// TwinCAT 3 PLC project SPS
// ProgramVersion: 3.1.4023.0
// libraries:
//   Tc2_MC2, * (Beckhoff Automation GmbH)
//   Tc2_NCI, * (Beckhoff Automation GmbH)
//   Tc2_PlcInterpolation, * (Beckhoff Automation GmbH)
//   Tc2_Standard, * (Beckhoff Automation GmbH)
//   Tc2_System, * (Beckhoff Automation GmbH)
//   Tc3_Module, * (Beckhoff Automation GmbH)
//   VisuDialogs, * (System)
//   VisuSymbols,3.5.10.0,System
// project tree:
//   DUTs/ E_AxesCmd.TcDUT, E_ButtonState.TcDUT, E_CheckMagazines_New.TcDUT, E_ErrorIDs.TcDUT, E_ErrorSrcs.TcDUT, E_GripperState.TcDUT, E_JobType.TcDUT, E_NC_State.TcDUT, E_NCI_State.TcDUT, E_PortalState.TcDUT, E_PortalState_New.TcDUT, E_ResetHW.TcDUT, E_SetJobState.TcDUT, ST_DeviceState.TcDUT, ST_Channel.TcDUT, ST_Light.TcDUT, ST_Error.TcDUT, ST_PortalJob.TcDUT, ST_PositionCmd.TcDUT, ST_SoftKey.TcDUT
//   / GlobalTextList.TcGTLO, PlcTask.TcTTO, Visualization Manager.TcVMO (not stored), VISU_TASK.TcTTO
//   GVLs/ HMI.TcGVL, GVL_CONST.TcGVL
//   POUs/Aktorik/ FB_AxesEnable.TcPOU, FB_AxisCtrl.TcPOU (excluded from build), FB_Gripper.TcPOU, FB_NciCtrl.TcPOU, FB_SimpleNcControl.TcPOU (excluded from build), FB_VI_Light.TcPOU
//   POUs/ FB_ErrorCollector.TcPOU, FB_IgorCtrl.TcPOU, FB_Portal.TcPOU, MAIN.TcPOU
//   POUs/Safety/ FB_SafeEStop.TcPOU, FB_SafeGroup.TcPOU, FB_SafeMon.TcPOU, FB_SafetyMonitoring.TcPOU
//   POUs/Zeug/ FB_BlockEconomySmart.TcPOU, FB_Error.TcPOU, FB_FuseControl.TcPOU, FB_FuseControl_1.TcPOU, I_NC_Ctrl.TcIO
//   VISUs/ VISU.TcVIS
// real-time tasks:
//   TASK PlcTask: cycle T#10ms, priority 20, ADS port 350
//   TASK PlcTask1: cycle T#10ms, priority 21, ADS port 351
//   TASK VISU_TASK: cycle T#50000us, priority 30, ADS port 352
// motion (NC):
//   TASK NC-Task 1 SAF: cycle T#2ms, priority 4, ADS port 501
//   TASK NC-Task 1 SVB: cycle T#10ms, priority 8, ADS port 511
//   AXIS X (id 1)
//     Dynamic: Acceleration=7500, Deceleration=7500, Jerk=20000, ToleranceBallAuxAxis=20
//     Velo: RefSearch=7.60333333333333, RefSync=7.60333333333333, SlowManual=38.0166666666667, FastManual=750, Fast=760.333333333333, Maximum=760.333
//     TargetPosControl: Range=0.5
//     PEHControl: Enable=true, Time=10
//     OtherSettings: AllowMotionCmdToSlave=true
//     encoder EncType=19
//       EncPara: ScaleFactorNumerator=20, ScaleFactorDenominator=1048576, Offset=150.930252075195, MaxCount=#xffffffff, ReferenceSystem=1
//         SoftEndMinControl: Enable=true, Range=-100
//         SoftEndMaxControl: Enable=true, Range=415
//         TimeComp: TimeCompMode=1
//     drive DrvType=16
//       DrvPara: MaxCount=#xffffffff, DriveControlDWord=#x00020100
//         Analog: VeloReferenz=836.366666666667, VeloScale=32, TorqueSetpointScale=10, ScaleFactorActTorque=0.004
//         TimeComp: TimeCompMode=1, TaskDelayCycles=1
//     controller CtrType=1
//       CtrPara: PriorControlFactor=1
//         PID: PosKp=30
//         Observer: BandWidth=20
//   AXIS Y (id 2)
//     Dynamic: Acceleration=2027.55, Deceleration=2027.55, Jerk=5406.81, ToleranceBallAuxAxis=20
//     Velo: RefSearch=7.60333333333333, RefSync=7.60333333333333, SlowManual=38.0166666666667, FastManual=700, Fast=760.333333333333, Maximum=760.333
//     TargetPosControl: Range=0.5
//     PEHControl: Enable=true, Time=10
//     OtherSettings: AllowMotionCmdToSlave=true
//     encoder EncType=19
//       EncPara: ScaleFactorNumerator=20, ScaleFactorDenominator=1048576, Offset=-52.5408172607422, MaxCount=#xffffffff, ReferenceSystem=1
//         SoftEndMinControl: Enable=true, Range=-2
//         SoftEndMaxControl: Enable=true, Range=300
//         TimeComp: TimeCompMode=1
//     drive DrvType=16
//       DrvPara: MaxCount=#xffffffff, DriveControlDWord=#x00020100
//         Analog: VeloReferenz=836.366666666667, VeloScale=32, TorqueSetpointScale=10, ScaleFactorActTorque=0.1
//         TimeComp: TimeCompMode=1, TaskDelayCycles=1
//     controller CtrType=1
//       CtrPara: PriorControlFactor=1
//         Observer: BandWidth=20
//   AXIS Z (id 3)
//     Dynamic: Acceleration=7500, Deceleration=7500, Jerk=20000, ToleranceBallAuxAxis=20
//     Velo: RefSearch=2.875, RefSync=2.875, SlowManual=14.375, FastManual=200.25, Fast=287.5, Maximum=287.5
//     TargetPosControl: Range=0.5
//     OtherSettings: AllowMotionCmdToSlave=true
//     encoder EncType=19
//       EncPara: ScaleFactorNumerator=5, ScaleFactorDenominator=1048576, Offset=69.1336441040039, Inverse=true, MaxCount=#xffffffff, ReferenceSystem=1
//         SoftEndMinControl: Enable=true
//         SoftEndMaxControl: Enable=true, Range=90
//         TimeComp: TimeCompMode=1
//     drive DrvType=16
//       DrvPara: Inverse=true, MaxCount=#xffffffff, DriveControlDWord=#x00020100
//         Analog: VeloReferenz=316.25, VeloScale=32, TorqueSetpointScale=10, ScaleFactorActTorque=0.1
//         TimeComp: TimeCompMode=1, TaskDelayCycles=1
//     controller CtrType=1
//       CtrPara: PriorControlFactor=1
//         PosDiffControl: Range=0.2
//         PID: PosKp=40
//         Observer: BandWidth=20
// I/O:
//   DEVICE Device, AmsNetId 192.168.1.150.4.1
//     +S1-BC1 (EK1100) [EK1100 EtherCAT Coupler (2A E-Bus)]
//       +S1-SI1 (EL1918) [EL1918, 8Ch. Safety Input 24V, TwinSAFE]
//         modules: Module 2 (FSLOGIC)
//       +S1-SO1 (EL2904) [EL2904, 4 Ch. Safety Output 24V, 0.5A, TwinSAFE]
//         modules: Module 1 (FSOES), Module 2 (DO)
//       +S1-DI1 (EL1804) [EL1804 4Ch. Dig. Input 24V, 3ms]
//       +S1-DI2 (EL1804) [EL1804 4Ch. Dig. Input 24V, 3ms]
//       +S1-DO1 (EL2004) [EL2004 4Ch. Dig. Output 24V, 0.5A]
//       +S1-PM1 (EL7211-9014) [EL7211-9014 1Ch. MDP742 Servo motor output stage with OCT (50V, 4.5A RMS) and STO input]
//       +S1-PM2 (EL7211-9014) [EL7211-9014 1Ch. MDP742 Servo motor output stage with OCT (50V, 4.5A RMS) and STO input]
//       +S1-PM3 (EL7211-9014) [EL7211-9014 1Ch. MDP742 Servo motor output stage with OCT (50V, 4.5A RMS) and STO input]
//       Term 20 (EK1310)
//     Box 21 (VIP2000-1010)
// variable links:
//   Device <-> Device/+S1-BC1 (EK1100)/+S1-SI1 (EL1918)
//     +S1-BC1 (EK1100)/+S1-SO1 (EL2904)/Module 1 (FSOES)/RxPDO/FSOE <-> ConnectionInputs/Message_13 TxPDO
//     +S1-BC1 (EK1100)/+S1-SO1 (EL2904)/Module 1 (FSOES)/TxPDO/FSOE <-> ConnectionOutputs/Message_13 RxPDO
//   NC-Task 1 SAF/Axes/X <-> Device/+S1-BC1 (EK1100)/+S1-PM1 (EL7211-9014)
//     Drive/Inputs/In/nDataIn1 <-> DRV Following error actual value/Following error actual value
//     Drive/Inputs/In/nDataIn3[0] <-> DRV Torque actual value/Torque actual value
//     Drive/Inputs/In/nDcOutputTime <-> InfoData/DcOutputShift
//     Drive/Inputs/In/nState1 <-> DRV Statusword/Statusword
//     Drive/Inputs/In/nState2 <-> DRV Statusword/Statusword @bit 8
//     Drive/Inputs/In/nState4 @bit 1 <-> WcState/InputToggle
//     Drive/Inputs/In/nState4 <-> WcState/WcState
//     Drive/Outputs/Out/nCtrl1 <-> DRV Controlword/Controlword
//     Drive/Outputs/Out/nCtrl2 <-> DRV Controlword/Controlword @bit 8
//     Drive/Outputs/Out/nDataOut1 <-> DRV Target position/Target position
//     Enc/Inputs/In/nDataIn1 <-> FB Position/Position
//     Enc/Inputs/In/nDcInputTime <-> InfoData/DcInputShift
//     Enc/Inputs/In/nState4 @bit 1 <-> WcState/InputToggle
//     Enc/Inputs/In/nState4 <-> WcState/WcState
//   NC-Task 1 SAF/Axes/Y <-> Device/+S1-BC1 (EK1100)/+S1-PM2 (EL7211-9014)
//     Drive/Inputs/In/nDataIn1 <-> DRV Following error actual value/Following error actual value
//     Drive/Inputs/In/nDcOutputTime <-> InfoData/DcOutputShift
//     Drive/Inputs/In/nState1 <-> DRV Statusword/Statusword
//     Drive/Inputs/In/nState2 <-> DRV Statusword/Statusword @bit 8
//     Drive/Inputs/In/nState4 @bit 1 <-> WcState/InputToggle
//     Drive/Inputs/In/nState4 <-> WcState/WcState
//     Drive/Outputs/Out/nCtrl1 <-> DRV Controlword/Controlword
//     Drive/Outputs/Out/nCtrl2 <-> DRV Controlword/Controlword @bit 8
//     Drive/Outputs/Out/nDataOut1 <-> DRV Target position/Target position
//     Enc/Inputs/In/nDataIn1 <-> FB Position/Position
//     Enc/Inputs/In/nDcInputTime <-> InfoData/DcInputShift
//     Enc/Inputs/In/nState4 @bit 1 <-> WcState/InputToggle
//     Enc/Inputs/In/nState4 <-> WcState/WcState
//   NC-Task 1 SAF/Axes/Z <-> Device/+S1-BC1 (EK1100)/+S1-PM3 (EL7211-9014)
//     Drive/Inputs/In/nDataIn1 <-> DRV Following error actual value/Following error actual value
//     Drive/Inputs/In/nDcOutputTime <-> InfoData/DcOutputShift
//     Drive/Inputs/In/nState1 <-> DRV Statusword/Statusword
//     Drive/Inputs/In/nState2 <-> DRV Statusword/Statusword @bit 8
//     Drive/Inputs/In/nState4 @bit 1 <-> WcState/InputToggle
//     Drive/Inputs/In/nState4 <-> WcState/WcState
//     Drive/Outputs/Out/nCtrl1 <-> DRV Controlword/Controlword
//     Drive/Outputs/Out/nCtrl2 <-> DRV Controlword/Controlword @bit 8
//     Drive/Outputs/Out/nDataOut1 <-> DRV Target position/Target position
//     Enc/Inputs/In/nDataIn1 <-> FB Position/Position
//     Enc/Inputs/In/nDcInputTime <-> InfoData/DcInputShift
//     Enc/Inputs/In/nState4 @bit 1 <-> WcState/InputToggle
//     Enc/Inputs/In/nState4 <-> WcState/WcState
//   SPS/SPS Instance <-> Device/+S1-BC1 (EK1100)/+S1-DI1 (EL1804)
//     PlcTask Inputs/MAIN.fbIgorCtrl.fbFuseControl.fbBlockFuse.In <-> Channel 3/Input
//     PlcTask Inputs/MAIN.fbIgorCtrl.fbFuseControl48V.bInFuse <-> Channel 4/Input
//     PlcTask Inputs/MAIN.fbIgorCtrl.fbPortal.fbGripper.bGripperFullClosed <-> Channel 2/Input
//     PlcTask Inputs/MAIN.fbIgorCtrl.fbPortal.fbGripper.bPartSensor <-> Channel 1/Input
//   SPS/SPS Instance <-> Device/+S1-BC1 (EK1100)/+S1-DI2 (EL1804)
//     PlcTask Inputs/MAIN.fbIgorCtrl.fbPortal.bStampZAxis <-> Channel 1/Input
//   SPS/SPS Instance <-> Device/+S1-BC1 (EK1100)/+S1-DO1 (EL2004)
//     PlcTask Outputs/MAIN.fbIgorCtrl.fbFuseControl.fbBlockFuse.Out <-> Channel 3/Output
//     PlcTask Outputs/MAIN.fbIgorCtrl.fbFuseControl48V.bOutFuse <-> Channel 4/Output
//     PlcTask Outputs/MAIN.fbIgorCtrl.fbPortal.fbGripper.bCloseGripper <-> Channel 2/Output
//     PlcTask Outputs/MAIN.fbIgorCtrl.fbPortal.fbGripper.bOpenGripper <-> Channel 1/Output
//   SPS/SPS Instance <-> Device/+S1-BC1 (EK1100)/+S1-PM1 (EL7211-9014)
//     PlcTask Inputs/MAIN.fbIgorCtrl.fbSafetyMonitoring.nDrvInfoData1 <-> DRV Info data 1/Info data 1
//   SPS/SPS Instance <-> Device/+S1-BC1 (EK1100)/+S1-PM2 (EL7211-9014)
//     PlcTask Inputs/MAIN.fbIgorCtrl.fbSafetyMonitoring.nDrvInfoData2 <-> DRV Info data 1/Info data 1
//   SPS/SPS Instance <-> Device/+S1-BC1 (EK1100)/+S1-PM3 (EL7211-9014)
//     PlcTask Inputs/MAIN.fbIgorCtrl.fbSafetyMonitoring.nDrvInfoData3 <-> DRV Info data 1/Info data 1
//   SPS/SPS Instance <-> Device/+S1-BC1 (EK1100)/+S1-SI1 (EL1918)
//     PlcTask Inputs/MAIN.fbIgorCtrl.fbPortal.bSafetyOK <-> StandardInputs/Standard Out Var 20
//     PlcTask Inputs/MAIN.fbIgorCtrl.fbSafetyMonitoring.bEStopButtonOk <-> StandardInputs/Standard Out Var 16
//     PlcTask Inputs/MAIN.fbIgorCtrl.fbSafetyMonitoring.bLightCurtainOk <-> StandardInputs/Standard Out Var 19
//     PlcTask Inputs/MAIN.fbIgorCtrl.fbSafetyMonitoring.fbEStop.nDiag <-> Function Block Info Data/SafetyGruppe.SafetyNetzwerk.FBEstop1 Info Data/Diag
//     PlcTask Inputs/MAIN.fbIgorCtrl.fbSafetyMonitoring.fbEStop.nState <-> Function Block Info Data/SafetyGruppe.SafetyNetzwerk.FBEstop1 Info Data/State
//     PlcTask Inputs/MAIN.fbIgorCtrl.fbSafetyMonitoring.fbGroup.nDiag <-> TwinSAFE Group Info Data/SafetyGruppe Info Data/Diag
//     PlcTask Inputs/MAIN.fbIgorCtrl.fbSafetyMonitoring.fbGroup.nState <-> TwinSAFE Group Info Data/SafetyGruppe Info Data/State
//     PlcTask Inputs/MAIN.fbIgorCtrl.fbSafetyMonitoring.fbMonEStop.nDiag <-> Function Block Info Data/SafetyGruppe.SafetyNetzwerk.FBMon1 Info Data/Diag
//     PlcTask Inputs/MAIN.fbIgorCtrl.fbSafetyMonitoring.fbMonEStop.nState <-> Function Block Info Data/SafetyGruppe.SafetyNetzwerk.FBMon1 Info Data/State
//     PlcTask Inputs/MAIN.fbIgorCtrl.fbSafetyMonitoring.fbMonLightCurtain.nDiag <-> Function Block Info Data/SafetyGruppe.SafetyNetzwerk.FBMon2 Info Data/Diag
//     PlcTask Inputs/MAIN.fbIgorCtrl.fbSafetyMonitoring.fbMonLightCurtain.nState <-> Function Block Info Data/SafetyGruppe.SafetyNetzwerk.FBMon2 Info Data/State
//     PlcTask Inputs/MAIN.fbIgorCtrl.fbSafetyMonitoring.fbMonSafetyGroup.nDiag <-> Function Block Info Data/SafetyGruppe.SafetyNetzwerk.FBMon3 Info Data/Diag
//     PlcTask Inputs/MAIN.fbIgorCtrl.fbSafetyMonitoring.fbMonSafetyGroup.nState <-> Function Block Info Data/SafetyGruppe.SafetyNetzwerk.FBMon3 Info Data/State
//     PlcTask Outputs/MAIN.fbIgorCtrl.fbPortal.bQuitEStop <-> StandardOutputs/Standard In Var 17
//     PlcTask Outputs/MAIN.fbIgorCtrl.fbPortal.bSafetyErrAck <-> StandardOutputs/Standard In Var 23
//     PlcTask Outputs/MAIN.fbIgorCtrl.fbPortal.bSafetyRun <-> StandardOutputs/Standard In Var 22
//     PlcTask Outputs/MAIN.fbIgorCtrl.fbSafetyMonitoring.bCollectEDM <-> StandardOutputs/Standard In Var 24
//   SPS/SPS Instance <-> Device/Box 21 (VIP2000-1010)
//     PlcTask Inputs/MAIN.fbIgorCtrl.fbLight.stDeviceState.Diag <-> Device/Main Inputs/Diag
//     PlcTask Inputs/MAIN.fbIgorCtrl.fbLight.stDeviceState.Error <-> Device/Main Inputs/Error
//     PlcTask Inputs/MAIN.fbIgorCtrl.fbLight.stDeviceState.Ready <-> Device/Main Inputs/Ready
//     PlcTask Inputs/MAIN.fbIgorCtrl.fbLight.stDeviceState.State <-> Device/Main Inputs/Status
//     PlcTask Inputs/MAIN.fbIgorCtrl.fbLight.stDeviceState.SwitchOnCnt <-> Device/Main Inputs/Switch-on counter
//     PlcTask Inputs/MAIN.fbIgorCtrl.fbLight.stDeviceState.Warning <-> Device/Main Inputs/Warning
//     PlcTask Inputs/MAIN.fbIgorCtrl.fbLight.stLight.bLightOn <-> Device/Opmode Continuous Inputs/Light on
//     PlcTask Outputs/MAIN.fbIgorCtrl.fbLight.stLight.bActive <-> Device/Opmode Continuous Outputs/Output
//     PlcTask Outputs/MAIN.fbIgorCtrl.fbLight.stLight.bEnable <-> Device/Main Outputs/Enable
//     PlcTask Outputs/MAIN.fbIgorCtrl.fbLight.stLight.bReset <-> Device/Main Outputs/Reset
//     PlcTask Outputs/MAIN.fbIgorCtrl.fbLight.stLight.channel[1]/bActive <-> Channel Red/ChContinuous Outputs/Active
//     PlcTask Outputs/MAIN.fbIgorCtrl.fbLight.stLight.channel[1]/nBrightness <-> Channel Red/ChContinuous Outputs/Brightness
//     PlcTask Outputs/MAIN.fbIgorCtrl.fbLight.stLight.channel[2]/bActive <-> Channel Blue/ChContinuous Outputs/Active
//     PlcTask Outputs/MAIN.fbIgorCtrl.fbLight.stLight.channel[2]/nBrightness <-> Channel Blue/ChContinuous Outputs/Brightness
//     PlcTask Outputs/MAIN.fbIgorCtrl.fbLight.stLight.channel[3]/bActive <-> Channel Green/ChContinuous Outputs/Active
//     PlcTask Outputs/MAIN.fbIgorCtrl.fbLight.stLight.channel[3]/nBrightness <-> Channel Green/ChContinuous Outputs/Brightness
//     PlcTask Outputs/MAIN.fbIgorCtrl.fbLight.stLight.channel[4]/bActive <-> Channel Orange/ChContinuous Outputs/Active
//     PlcTask Outputs/MAIN.fbIgorCtrl.fbLight.stLight.channel[4]/nBrightness <-> Channel Orange/ChContinuous Outputs/Brightness
//   SPS/SPS Instance <-> NC-Task 1 SAF/Axes/X
//     PlcTask Inputs/MAIN.fbIgorCtrl.fbPortal.aAxis[0].NcToPlc <-> Outputs/ToPlc
//     PlcTask Outputs/MAIN.fbIgorCtrl.fbPortal.aAxis[0].PlcToNc <-> Inputs/FromPlc
//   SPS/SPS Instance <-> NC-Task 1 SAF/Axes/Y
//     PlcTask Inputs/MAIN.fbIgorCtrl.fbPortal.aAxis[1].NcToPlc <-> Outputs/ToPlc
//     PlcTask Outputs/MAIN.fbIgorCtrl.fbPortal.aAxis[1].PlcToNc <-> Inputs/FromPlc
//   SPS/SPS Instance <-> NC-Task 1 SAF/Axes/Z
//     PlcTask Inputs/MAIN.fbIgorCtrl.fbPortal.aAxis[2].NcToPlc <-> Outputs/ToPlc
//     PlcTask Outputs/MAIN.fbIgorCtrl.fbPortal.aAxis[2].PlcToNc <-> Inputs/FromPlc
//   SPS/SPS Instance <-> NC-Task 1 SAF/Interpolation Channel
//     PlcTask Inputs/MAIN.fbIgorCtrl.fbPortal.fbNciCtrl.stItpToPlc <-> Outputs/ToPlc
//     PlcTask Outputs/MAIN.fbIgorCtrl.fbPortal.fbNciCtrl.stPlcToItp <-> Inputs/FromPlc

CONFIGURATION SPS
    RESOURCE PLC ON TwinCAT3
        TASK PlcTask(INTERVAL := T#10ms, PRIORITY := 21);
        TASK VISU_TASK(INTERVAL := T#50000us, PRIORITY := 30);
        PROGRAM MAIN WITH PlcTask : MAIN;
        PROGRAM VisuElems_Visu_Prg WITH VISU_TASK : VisuElems.Visu_Prg;
    END_RESOURCE
END_CONFIGURATION

// ---- DUTs/E_AxesCmd.TcDUT
TYPE E_AxesCmd :
(
	E_AxesCmd_IDLE := 0,
	E_AxesCmd_RESET := 10,
	E_AxesCmd_MOVE_ABS := 20,
	E_AxesCmd_MOVE_REL := 30,
	E_AxesCmd_JOG := 40,
	E_AxesCmd_REFERENCING := 50,
	E_AxesCmd_STOP := 70,
	E_AxesCmd_FINISHED := 80,
	E_AxesCmd_ERROR := 99
);
END_TYPE

// ---- DUTs/E_ButtonState.TcDUT
{attribute 'strict'}
TYPE E_ButtonState :
(
	E_ButtonState_OFF := 0,
	E_ButtonState_ON,
	E_ButtonState_BLINK
);
END_TYPE

// ---- DUTs/E_CheckMagazines_New.TcDUT
{attribute 'qualified_only'}
{attribute 'strict'}
TYPE E_CheckMagazines_New :
(
	eIdle	:= 0,
	eStartNewNCI	:= 1,
	eDebug := 2,
	eWaitForPortal := 3
);
END_TYPE

// ---- DUTs/E_ErrorIDs.TcDUT
{attribute 'qualified_only'}
{attribute 'strict'}
TYPE E_ErrorIDs :
(
	eNoError := 0,
	eUndefinedError := 1,
	eUndefinedState := 2,
	
	eInvalidReference := 21,
	
	eAxisRelease := 31,
	eAbsMove := 32,
	eRelMove := 33,
	eJog := 34,
	eStopAxis := 35,
	eResetAxis := 36,
	eAxesNotReady := 37,
	eAxisError := 38,
	
	eTimeout := 41,
	eInvalidData := 42,
	eReset := 43,
	
	eBuildGroup := 51,
	eClearGroup := 52,
	eFillTable := 53,
	eNotAllowedDriveDown := 54,
	
	eSafetyFbError := 61,
	eCommError := 62,
	eModuleFault := 63,
	eCompareError := 64,
	eEStopPressed := 65,
	eLightCurtain := 66,
	
	eNoStoneInGripper := 71,
	eMagEmpty := 72,
	
	eFuseTripped := 81,
	eFuseOff := 82,
	eFuseOvercurrent := 83,
	
	eClearFieldNoCapacityFound := 90,
	eNoJobsFound := 91,
	eStamp := 92,
	eNoStonesFound := 93,
	
	eCtrlOff := 99
);
END_TYPE

// ---- DUTs/E_ErrorSrcs.TcDUT
{attribute 'qualified_only'}
{attribute 'strict'}
TYPE E_ErrorSrcs :
(
	eNoError := 0,
	ePlc := 1,
	eAxisX := 2,
	eAxisY := 3,
	eAxisZ := 4,
	eAxisGroup := 5,
	eAxisCtrlPtp := 6,
	eAxisCtrlNci := 7,
	eAxisCtrl := 8,
	eGripper := 9,
	eSafety := 10,
	eSafetyGroup := 11,
	eSafetyFb := 12,
	ePortal := 13,
	eFuse := 14
);
END_TYPE

// ---- DUTs/E_GripperState.TcDUT

TYPE E_GripperState :
(
	E_GripperState_INIT := 0,
	E_GripperState_OPENING,
	E_GripperState_OPENED,
	E_GripperState_CLOSING,
	E_GripperState_CLOSED,
	E_GripperState_UNDEFINED
);
END_TYPE

// ---- DUTs/E_JobType.TcDUT
TYPE E_JobType :
(
	E_JobType_MoveStone,
	E_JobType_NewStone,
	E_JobType_RemoveStone
);
END_TYPE

// ---- DUTs/E_NC_State.TcDUT
TYPE E_NC_State :
(
	E_NC_State_INIT := 0,
	E_NC_State_IDLE := 1,
	E_NC_State_RUN := 7,
	E_NC_State_ABORT := 8,
	E_NC_State_ERROR := 9
);
END_TYPE

// ---- DUTs/E_NCI_State.TcDUT
TYPE E_NCI_State :
(
	E_NCI_State_INIT := 0,
	E_NCI_State_IDLE := 1,
	E_NCI_State_BUILD_GROUP := 4,
	E_NCI_State_LOAD_CODE := 5,
	E_NCI_State_FEED_TABLE := 6,
	E_NCI_State_RUN := 7,
	E_NCI_State_ABORT := 8,
	E_NCI_State_CLEAR_GROUP := 9,
	E_NCI_State_ESTOP := 90,
	E_NCI_State_ERROR := 99
);
END_TYPE

// ---- DUTs/E_PortalState.TcDUT
TYPE E_PortalState :
(
	E_PortalState_INIT := 0,
	E_PortalState_IDLE,
	E_PortalState_SET_JOB,
	E_PortalState_MOVE_TO_STONE,
	E_PortalState_TRANSPORT_STONE,
	E_PortalState_WAITGRIPPER_OPEN,
	E_PortalState_WAITGRIPPER_CLOSE,
	E_PortalState_HOME,
	E_PortalState_ESTOP,
	E_PortalState_AFTER_ESTOP,
	E_PortalState_MANUAL_MODE,
	E_PortalState_SCAN_MAGS,
	E_PortalState_ERROR := 99
);
END_TYPE

// ---- DUTs/E_PortalState_New.TcDUT
TYPE E_PortalState_New :
(
	eInit := 0,
	eIdle,
	eSetJob,
	eOpenGripper,
	eCloseGripper,
	eError,
	eMoveToStone,
	eTrspStone,
	eStampTriggered,
	eHome,
	eEStop,
	eAfterEStop,
	eManualMode,
	eDebug
);
END_TYPE

// ---- DUTs/E_ResetHW.TcDUT
{attribute 'qualified_only'}
{attribute 'strict'}
TYPE E_ResetHW :
(
	INIT := 0,
	RESET_HW := 10,
	DONE := 50
);
END_TYPE

// ---- DUTs/E_SetJobState.TcDUT
{attribute 'qualified_only'}
{attribute 'strict'}
TYPE E_SetJobState :
(
	eIdle := 0,
	eAxesNotReady,
	eSelNewStone,
	eSelRemoveStone,
	eCheckAllMagazines,
	eValidateNewStone,
	eValidateRemoveStone
);
END_TYPE

// ---- DUTs/ST_DeviceState.TcDUT
TYPE ST_DeviceState :
STRUCT
	Ready		AT%I*	: BIT;
	Warning		AT%I*	: BIT;
	Error		AT%I*	: BIT;
	Diag		AT%I*	: BIT;
	State		AT%I*	: UDINT;
	SwitchOnCnt	AT%I*	: UDINT;
END_STRUCT
END_TYPE

// ---- DUTs/ST_Channel.TcDUT
TYPE ST_Channel :
STRUCT
	bActive				AT %Q*  : BOOL	 := FALSE;	
	nBrightness			AT %Q*	: UINT	 := 100; 
END_STRUCT
END_TYPE

// ---- DUTs/ST_Light.TcDUT
TYPE ST_Light :
STRUCT
	bEnable					AT %Q* 	: BOOL := TRUE;				// Global enable of light
	bReset					AT %Q*	: BOOL := FALSE;			// Reset light
	bActive					AT %Q*  : BOOL	 := FALSE;			// General activation of the light, depends on the chanels
	bLightOn				AT %I*	: BOOL;						// Light is activated
	channel					AT %Q*  : ARRAY[1..4] OF ST_Channel; // 1: IR, 2: blue, 3: green, 4: orange
	nTemperature			AT %I*	: SINT;						// temperature channel
END_STRUCT
END_TYPE

// ---- DUTs/ST_Error.TcDUT
TYPE ST_Error :
STRUCT
	nSource:		UDINT;
	nType:			UDINT;
	sMsg:			STRING(80);
END_STRUCT
END_TYPE

// ---- DUTs/ST_PortalJob.TcDUT
TYPE ST_PortalJob :
STRUCT
	nJobID:			UDINT; //Job Nummer
	eJobType:		E_JobType;  //Neuer Stein von Stapel oder Stein auf Brett oder Stein entfernen
	fStartPosX:		LREAL; //Startposition x in mm
	fStartPosY:		LREAL; //Startposition y in mm
	fDestPosX:		LREAL; //Zielposition x in mm
	fDestPosY:		LREAL; //Zielposition y in mm
	bBlack:			BOOL; //entscheidet über Lagerposition
END_STRUCT
END_TYPE

// ---- DUTs/ST_PositionCmd.TcDUT
TYPE ST_PositionCmd :
STRUCT
	nNo:	UDINT;
	fPosX:	LREAL;
	fPosY:	LREAL;
	fPosZ:	LREAL;
	fVelo:	LREAL;
	bExact:	BOOL;
END_STRUCT
END_TYPE

// ---- DUTs/ST_SoftKey.TcDUT
TYPE ST_SoftKey :
STRUCT
	bIsPressed:	BOOL;
	eState:		E_ButtonState;
END_STRUCT
END_TYPE

// ---- GVLs/HMI.TcGVL
{attribute 'qualified_only'}
VAR_GLOBAL	
//TO HMI
	bErrorChange:		BOOL;
	aErrors:			ARRAY [0..MAX_ERRORS - 1] OF ST_Error;
	nNumberErrors:		UINT;
	bSafetyOK:			BOOL;
	bPortalBusy:		BOOL;
	bInManual:			BOOL;
	bGripperOpen:		BOOL;
	bGripperClosed:		BOOL;
	bHandInPortal:		BOOL; 
	
//FROM HMI
	bQuit:				BOOL;
	
	bSetJob:			BOOL;
	stJob:				ST_PortalJob;
	stLastJob:			ST_PortalJob;
     	
	bReqManualCtrl:		BOOL := TRUE;
	bOpenGripper:		BOOL;
	bCloseGripper:		BOOL;
	bSafetyRun:			BOOL;
	
	bLightOn:			BOOL;
	bLightWin: 			BOOL;
	bLightLose:			BOOL;
	
	bLightParty: 		BOOL;
	
	bAllJobsSend: 		BOOL; 
	
//TO AND FROM HMI
	stSoftKeyCtrlOn:	ST_SoftKey;
	stSoftKeyCtrlOff:	ST_SoftKey;
	stSoftKeyAutoOn:	ST_SoftKey;
	stSoftKeyAutoOff:	ST_SoftKey;
	stSoftKeyQuit:		ST_SoftKey;

//system
	fbErrorCollector:	FB_ErrorCollector;
	
//parameters
	fAxesOverride:		LREAL := 100.0;
	fAxesOverrideMan:	LREAL := 20.0;
	
	fPortalPosIdleX:	LREAL := -20;
	fPortalPosIdleY:	LREAL := 0;
	fPortalPosIdleZ:	LREAL := 50;

	fScreenPosOffsetX:	LREAL := 0;
	fScreenPosOffsetY:	LREAL := 0;
END_VAR

// ---- GVLs/GVL_CONST.TcGVL
VAR_GLOBAL CONSTANT	
	STONE_POS_FIELD_Z:	LREAL := 1;
	MIN_MOVE_HEIGHT_Z:	LREAL := 40; //beachte: Stäbe von Magazin ca. 35 mm -> nicht unter 40 stellen!
	STONE_HEIGHT:		LREAL := 8; //Steinhöhe in mm -> für Positionen in Magazin
	
	MAX_JOB_COUNT:		USINT := 30;
	MAX_ERRORS:			USINT := 55;
	
	X:					USINT := 0;
	Y:					USINT := 1;
	Z:					USINT := 2;
	
	MAGAZINE_NUMBER:	USINT := 6; //Anzahl Magazine
	MAGAZINE_CAPACITY:	USINT := 4;	//Anzahl Positionen pro Magazin	
	
(******Stapel für Spielsteine******)
	STACK_POS_X:			LREAL := -97.2; 
	STACK_1_POS_Y:			LREAL := 52.6;	
	STACK_2_POS_Y:			LREAL := STACK_1_POS_Y + 28;
	STACK_3_POS_Y:			LREAL := STACK_2_POS_Y + 28;
	STACK_4_POS_Y:			LREAL := STACK_3_POS_Y + 94;
	STACK_5_POS_Y:			LREAL := STACK_4_POS_Y + 28;
	STACK_6_POS_Y:			LREAL := STACK_5_POS_Y + 28;//258.6
	STACK_POS_Z_BASE:		LREAL := 3;
	STACK_POS_Z_BASE_REMOVE:LREAL := 8;
	
(******Positionen Magazin-Scan******)
	STACK_SCAN_POS_X:		LREAL := -59;
	STACK_1_SCAN_POS_Y:		LREAL := STACK_1_POS_Y + 33.8;
	STACK_2_SCAN_POS_Y:		LREAL := STACK_2_POS_Y + 33.8;
	STACK_3_SCAN_POS_Y:		LREAL := STACK_3_POS_Y + 33.8;
	STACK_4_SCAN_POS_Y:		LREAL := STACK_4_POS_Y + 33.8;
	STACK_5_SCAN_POS_Y:		LREAL := STACK_5_POS_Y + 33.8;
	STACK_6_SCAN_POS_Y:		LREAL := STACK_6_POS_Y + 33.8;
	STACK_SCAN_POS_Z_BASE:	LREAL := 8.5;
	
END_VAR

// ---- POUs/Zeug/I_NC_Ctrl.TcIO
INTERFACE I_NC_Ctrl

METHOD M_AxisRef
VAR_INPUT
	rX:		REFERENCE TO AXIS_REF;
	rY:		REFERENCE TO AXIS_REF;
	rZ:		REFERENCE TO AXIS_REF;
END_VAR
END_METHOD

METHOD M_CancleJob
VAR_INPUT
END_VAR
END_METHOD

METHOD M_Cyclic
VAR_INPUT
END_VAR
END_METHOD

METHOD M_NewJob
VAR_INPUT
	fTargetPosX:	LREAL;
	fTargetPosY:	LREAL;
	fTargetPosZ:	LREAL;
END_VAR
END_METHOD

PROPERTY P_bInductiveSensor : BOOL
SET
END_SET
END_PROPERTY

PROPERTY P_Busy : BOOL
GET
END_GET
END_PROPERTY

PROPERTY P_Enable : BOOL
SET
END_SET
END_PROPERTY

PROPERTY P_ErrID : E_ErrorIDs
GET
END_GET
END_PROPERTY

PROPERTY P_Error : BOOL
GET
END_GET
END_PROPERTY

PROPERTY P_ErrSrc : E_ErrorSrcs
GET
END_GET
END_PROPERTY

PROPERTY P_ReadyForJob : BOOL
GET
END_GET
END_PROPERTY

PROPERTY P_Reset : BOOL
SET
END_SET
END_PROPERTY

END_INTERFACE

// ---- POUs/MAIN.TcPOU
PROGRAM MAIN
VAR
	fbIgorCtrl:			FB_IgorCtrl;
END_VAR

fbIgorCtrl();

END_PROGRAM

// ---- POUs/FB_IgorCtrl.TcPOU
FUNCTION_BLOCK FB_IgorCtrl
VAR_INPUT
END_VAR
VAR_OUTPUT
	fbError:	FB_Error;
END_VAR
VAR
	fbPortal:			FB_Portal;
	fbSafetyMonitoring:	FB_SafetyMonitoring;
	fbFuseControl:		FB_FuseControl;
	fbFuseControl48V: 	FB_FuseControl_1;
	fbLight			:	FB_VI_Light;
END_VAR

VAR
	fbBlinkTimer1		: TON;
	fbBlinkTimer2		: TON;
	fbTimer				: TON;
	fbRS				: RS;
	nCntParty			: UINT;
	rTrig1				: R_TRIG;
	rTrig2				: R_TRIG;
	
	nRed				: UINT;
	nGreen				: UINT;
	nBlue				: UINT;
END_VAR

A_HmiComm();

fbSafetyMonitoring();

fbFuseControl();
fbFuseControl48V(bResetChannels := HMI.bQuit);


fbPortal(
	bFuseOk := NOT fbFuseControl.fbError.bError,
	bFuse48VOk := NOT fbFuseControl.fbError.bError,
	bManualMode:= HMI.bReqManualCtrl, 
	stNewJob:= HMI.stJob, 
	bImportJob:= HMI.bSetJob,
	bQuit:= HMI.bQuit OR fbPortal.bQuit,//kann quit nicht false setzen
	bSafetyRun := HMI.bSafetyRun,
	bSafetyOK=> HMI.bSafetyOK, 
	bBusy=> HMI.bPortalBusy,
	fbError=> );

HMI.bGripperClosed := fbPortal.fbGripper.bGripperClosed;
HMI.bGripperOpen := fbPortal.fbGripper.bGripperOpen;

IF NOT HMI.bSafetyRun AND NOT fbError.bError THEN
	fbError.M_Set(1, 'Steuerung ausgeschaltet', 0, E_ErrorIDs.eCtrlOff, E_ErrorSrcs.ePlc);
ELSIF HMI.bSafetyRun AND fbError.bError THEN
	fbError.M_Reset();
END_IF

//Set trigger white light
IF HMI.bLightOn THEN
	HMI.bLightWin := FALSE;
	HMI.bLightLose := FALSE;
	fbLight(bLightOn:= HMI.bLightOn);
	fbLight.bLightOn := FALSE;
	fbLight.SetIRGB(255, 255, 255, 255, 100);
ELSIF NOT HMI.bLightWin AND NOT HMI.bLightLose THEN
	fbLight(bLightOn:= HMI.bLightOn);
END_IF

//Set light for win
IF HMI.bLightWin AND NOT HMI.bLightLose AND NOT HMI.bLightOn THEN
	fbTimer(IN := TRUE, PT := T#3S);
	fbRS(SET := TRUE, RESET1 := fbTimer.Q);
	
	fbBlinkTimer1(IN := fbRS.Q1 AND NOT fbBlinkTimer2.Q, PT := T#0.5S, Q => fbLight.bLightOn);
	fbBlinkTimer2(IN := fbBlinkTimer1.Q, PT := T#0.5S);
	fbLight.SetIRGB(0, 0, 255, 0, 50);
	
	IF fbTimer.Q THEN
		HMI.bLightWin := FALSE;
		fbLight.bLightOn := FALSE;
		fbTimer(IN := FALSE);
		fbRS(SET := FALSE, RESET1 := TRUE);
	END_IF
	
	fbLight();
ELSE
	fbRS(SET := FALSE, RESET1 := FALSE);
END_IF

//set light for lose
IF HMI.bLightLose AND NOT HMI.bLightWin AND NOT HMI.bLightOn THEN
	fbTimer(IN := TRUE, PT := T#3S);
	fbRS(SET := TRUE, RESET1 := fbTimer.Q);
	
	fbBlinkTimer1(IN := fbRS.Q1 AND NOT fbBlinkTimer2.Q, PT := T#0.5S, Q => fbLight.bLightOn);
	fbBlinkTimer2(IN := fbBlinkTimer1.Q, PT := T#0.5S);
	fbLight.SetIRGB(0, 255, 0, 0, 50);
	
	IF fbTimer.Q THEN
		HMI.bLightLose := FALSE;
		fbLight.bLightOn := FALSE;
		fbTimer(IN := FALSE);
		fbRS(SET := FALSE, RESET1 := TRUE);
	END_IF
	
	fbLight();
ELSE
	fbRS(SET := FALSE, RESET1 := FALSE);
END_IF

//Party-Modus
IF HMI.bLightParty THEN
	fbTimer(IN := TRUE, PT := T#30S);
	fbRS(SET := TRUE, RESET1 := fbTimer.Q);
	
	fbBlinkTimer1(IN := fbRS.Q1 AND NOT fbBlinkTimer2.Q, PT := T#0.4S, Q => );
	fbBlinkTimer2(IN := fbBlinkTimer1.Q, PT := T#0.2S);
	fbLight.bLightOn := NOT fbBlinkTimer1.Q;
	IF rTrig1.Q OR rTrig2.Q THEN
		nCntParty := nCntParty + 1;
	END_IF
	
	CASE nCntParty OF 
		0: fbLight.SetIRGB(0, 255, 0, 0, 25);
		1: fbLight.SetIRGB(0, 255, 30, 0, 25);
		2: fbLight.SetIRGB(0, 255, 255, 0, 25);
		3: fbLight.SetIRGB(0, 180, 255, 0, 25);
		4: fbLight.SetIRGB(0, 0, 255, 0, 25);
		5: fbLight.SetIRGB(0, 0, 255, 150, 25);
		6: fbLight.SetIRGB(0, 0, 255, 255, 25);
		7: fbLight.SetIRGB(0, 0, 120, 255, 25);
		8: fbLight.SetIRGB(0, 0, 0, 255, 25);
		9: fbLight.SetIRGB(0, 120, 0, 255, 25);
		10: fbLight.SetIRGB(0, 255, 0, 120, 25); nCntParty := 0;
	END_CASE

	IF fbTimer.Q THEN
		HMI.bLightParty := FALSE;
		nCntParty := 0;
		fbLight.bLightOn := FALSE;
		fbTimer(IN := FALSE);
		fbRS(SET := FALSE, RESET1 := TRUE);
	END_IF
	
	rTrig1(CLK := fbBlinkTimer1.Q);
	rTrig2(CLK := fbBlinkTimer2.Q);
	fbLight();
ELSE
	fbRS(SET := FALSE, RESET1 := FALSE);
END_IF

ACTION A_HmiComm:
IF HMI.stSoftKeyCtrlOn.bIsPressed THEN
	HMI.bSafetyRun := TRUE;
END_IF
IF HMI.stSoftKeyCtrlOff.bIsPressed THEN
	HMI.bSafetyRun := FALSE;
END_IF
IF HMI.stSoftKeyAutoOn.bIsPressed THEN
	HMI.bReqManualCtrl := FALSE;
END_IF
IF HMI.stSoftKeyAutoOff.bIsPressed THEN
	HMI.bReqManualCtrl := TRUE;
END_IF

HMI.bInManual := MAIN.fbIgorCtrl.fbPortal.ePortalState = E_PortalState_New.eManualMode;

HMI.bHandInPortal := NOT MAIN.fbIgorCtrl.fbSafetyMonitoring.bLightCurtainOk;

HMI.bQuit := HMI.stSoftKeyQuit.bIsPressed;

IF HMI.bSafetyOK THEN
	HMI.stSoftKeyCtrlOn.eState := E_ButtonState_ON;
	HMI.stSoftKeyCtrlOff.eState := E_ButtonState_OFF;
	
	IF HMI.bReqManualCtrl THEN
		IF Main.fbIgorCtrl.fbPortal.ePortalState <> E_PortalState_New.eManualMode THEN
			HMI.stSoftKeyAutoOn.eState := E_ButtonState_BLINK;
			HMI.stSoftKeyAutoOff.eState := E_ButtonState_OFF;
		ELSE
			HMI.stSoftKeyAutoOn.eState := E_ButtonState_OFF;
			HMI.stSoftKeyAutoOff.eState := E_ButtonState_ON;
		END_IF
	ELSE
		IF HMI.nNumberErrors = 0 THEN
			HMI.stSoftKeyAutoOn.eState := E_ButtonState_ON;
			HMI.stSoftKeyAutoOff.eState := E_ButtonState_OFF;
		ELSE
			HMI.stSoftKeyAutoOn.eState := E_ButtonState_OFF;
			HMI.stSoftKeyAutoOff.eState := E_ButtonState_BLINK;
		END_IF
	END_IF
	
	IF HMI.nNumberErrors > 0 THEN
		HMI.stSoftKeyQuit.eState := E_ButtonState_BLINK;
	ELSE
		HMI.stSoftKeyQuit.eState := E_ButtonState_OFF;
	END_IF
ELSE
	HMI.stSoftKeyAutoOn.eState := E_ButtonState_OFF;
	HMI.stSoftKeyAutoOff.eState := E_ButtonState_ON;
	IF HMI.bSafetyRun THEN
		HMI.stSoftKeyCtrlOn.eState := E_ButtonState_BLINK;
		HMI.stSoftKeyCtrlOff.eState := E_ButtonState_OFF;
		HMI.stSoftKeyQuit.eState := E_ButtonState_BLINK;
	ELSE
		HMI.stSoftKeyCtrlOn.eState := E_ButtonState_OFF;
		HMI.stSoftKeyCtrlOff.eState := E_ButtonState_ON;
		HMI.stSoftKeyQuit.eState := E_ButtonState_OFF;
	END_IF
END_IF
END_ACTION

END_FUNCTION_BLOCK

// ---- POUs/Zeug/FB_Error.TcPOU
{attribute 'reflection'}
FUNCTION_BLOCK FB_Error
VAR_OUTPUT
	bError:		BOOL;
	nErrorID:	UDINT;
	eErrorID:	E_ErrorIDs;
	eErrorSrc:	E_ErrorSrcs;
	sErrorMsg:	STRING(128);
	nState:		INT; //State in dem der Error aufgetreten ist
	
	//{attribute 'instance-path'}
	//{attribute 'no_init'}
	//sSource:	STRING;
END_VAR

METHOD M_Reset
VAR_INPUT
END_VAR
IF bError THEN
	HMI.fbErrorCollector.M_QuitError(eErrorID, eErrorSrc);
	MEMSET(ADR(THIS^), 0, SIZEOF(THIS^));
END_IF
END_METHOD

METHOD M_Set
VAR_INPUT
	nID:	UDINT;
	sMsg:	STRING;
	nState:	INT; //State in dem der Error aufgetreten ist
	eID:	E_ErrorIDs;
	eSrc:	E_ErrorSrcs;
END_VAR
VAR_INST
	
END_VAR
IF NOT bError THEN
	bError := TRUE;
	nErrorID := nID;
	sErrorMsg := sMsg;
	THIS^.nState := nState;
	eErrorID := eID;
	eErrorSrc := eSrc;
	HMI.fbErrorCollector.M_NewError(eID, eSrc, sMsg);
END_IF
END_METHOD

END_FUNCTION_BLOCK

// ---- POUs/FB_Portal.TcPOU
FUNCTION_BLOCK FB_Portal
VAR_INPUT
	bManualMode:			BOOL;	                    	
	stNewJob:				ST_PortalJob;
	bImportJob:				BOOL;
	bQuit:					BOOL;
	bFuseOk:				BOOL;
	bFuse48VOk:				BOOL;
	bSafetyRun AT %Q*:		BOOL;
END_VAR
VAR CONSTANT	
END_VAR                 	
VAR_OUTPUT          		
	bBusy:					BOOL;
	fbError:				FB_Error;
	                    	
	//Safety            	
	bSafetyOK AT %I*:		BOOL := TRUE;
END_VAR             		
VAR                     
	//Safety            	
	bQuitEStop AT %Q*:		BOOL;
	bSafetyErrAck AT %Q*:	BOOL;
	
	//Sensor Stempeln		
	bStampZAxis				AT %I*	: BOOL;
	rTrigStamp:				R_TRIG;
	bStampReset: 			BOOL;
	
	fbRTrigSafety:			R_TRIG;
	                    	
	ePortalState:			E_PortalState_New;
	eTargetPortalState: 	E_PortalState_New;
	                    	
	fbGripper:				FB_Gripper := (bEnable := TRUE);
  
	aAxis:					ARRAY [X..Z] OF AXIS_REF;
	fbAxesEnable:			FB_AxesEnable;
	fbResetAxis:			MC_Reset; 
	                    	
	ipNcCtrl:				I_NC_Ctrl;
	fbNciCtrl:				FB_NciCtrl;
	                    	
	bMagazineTrack:			BOOL; //Anzahl steine in Magazinen bekannt? false wenn Spieler eingreift oder nicht initialisiert
	                    	
	stActJob:				ST_PortalJob;
	aJobBuffer:				ARRAY [0..MAX_JOB_COUNT - 1] OF ST_PortalJob;
	nJobCount:				USINT;
	i, k:					USINT;
	                    	
	aMagCounter:			ARRAY [0..MAGAZINE_NUMBER-1] OF USINT; //Anzahl Steine in Magazinen
	aMagSkipCheck:			ARRAY [0..MAGAZINE_NUMBER-1] OF BOOL;
	aMagYPositions:			ARRAY [0..MAGAZINE_NUMBER-1] OF LREAL; //Mitte Y
	aMagYScanPositions:		ARRAY [0..MAGAZINE_NUMBER-1] OF LREAL;
	fStonePosZFromMag:		LREAL; //berechnete Z pos für Stein aus Magazin
	nMag:					INT;
	nSelectedMag:			INT;
	nPosInMag:				USINT;
	bValidateStonePos:		BOOL;
	nValidationValue:		INT;
	bLastJobBlack:			BOOL;
	
//MAG Check
	nStonesInMag:				INT := MAGAZINE_CAPACITY;
	bWaitPortal, bCheck:		BOOL;
	bCheckedAllMag: 	BOOL;
	nNumChecked:				INT;
	rTrigCheck:			R_TRIG;
//New
	nCntActiveJobs		: SINT;
	nCntRemoveStones	: SINT;
	eCheckMagState		: E_CheckMagazines_New;
	nStonesInMagazin	: USINT := MAGAZINE_CAPACITY;
	
	bAllJobsReceived	: BOOL;
	
	nStateJobSelect		: INT;
	
	bReady				: BOOL;
	
	fTrigNCIDone		: F_TRIG;
	
	fSetJobHeight	: LREAL;
	
	bNCIJobStarted : BOOL;
	
	eSetJobState	: E_SetJobState;
END_VAR

IF ipNcCtrl <> 0 THEN
	A_Cycle();
ELSIF ePortalState <> E_PortalState_INIT THEN
	fbError.M_Set(1, 'Interface nicht referenziert', ePortalState, E_ErrorIDs.eInvalidReference, E_ErrorSrcs.ePlc);
	RETURN;
END_IF
fTrigNCIDone(CLK := fbNciCtrl.P_Busy);

CASE ePortalState OF
	E_PortalState_New.eInit:
		A_Init();
		ePortalState := E_PortalState_New.eIdle;
		
	E_PortalState_New.eIdle:
		IF NOT bManualMode THEN
			IF aJobBuffer[0].nJobID <> 0 THEN
				fbAxesEnable.M_EnableAxes();
				IF fbGripper.bGripperOpen THEN
					IF HMI.bAllJobsSend THEN	
						nValidationValue := 0;	//TODO: entfernen wenn eSetJobState verwendet
						bReady := FALSE;
						nNumChecked := 0;		//TODO: entfernen wenn eSetJobState verwendet
						nStateJobSelect := 0;
						ePortalState := E_PortalState_New.eSetJob;
					END_IF
				ELSE
					eTargetPortalState := E_PortalState_New.eIdle;
					ePortalState := E_PortalState_New.eOpenGripper;
				END_IF
			END_IF
		ELSE	//Handbetrieb
			ipNcCtrl.P_Enable := FALSE;
			fbAxesEnable.M_EnableAxes();
			ePortalState := E_PortalState_New.eManualMode;
		END_IF
	
	E_PortalState_New.eOpenGripper:
		fbGripper(bEnable := TRUE, bOpen := TRUE, bClose := FALSE);
		IF NOT fbGripper.bBusy AND fbGripper.bGripperOpen THEN
			IF eTargetPortalState = E_PortalState_New.eIdle THEN
				fbGripper(bOpen := FALSE);
				ePortalState := eTargetPortalState;	
			ELSE
				IF NOT fbGripper.fbError.bError THEN
					IF stActJob.nJobID <> 0 THEN	//aktuellen Auftrag umgesetzt
						IF stActJob.eJobType = E_JobType.E_JobType_RemoveStone AND nCntActiveJobs = 1 THEN
							aMagCounter[nSelectedMag] := aMagCounter[nSelectedMag] + nCntRemoveStones;
							nCntRemoveStones := 0;
						END_IF
						nCntActiveJobs := nCntActiveJobs - 1;
						HMI.stLastJob := stActJob;
						A_DequeueJob();
						IF nCntActiveJobs <= 0 THEN
							bReady := FALSE;
						END_IF
					ELSE
						bReady := FALSE;
					END_IF
					IF nJobCount = 0 THEN
						ipNcCtrl.M_NewJob(HMI.fPortalPosIdleX, HMI.fPortalPosIdleY, HMI.fPortalPosIdleZ); //Auftrag zu Home-Pos
						ePortalState := E_PortalState_New.eHome;
					ELSE
						ePortalState := E_PortalState_New.eSetJob;	
					END_IF			
				ELSE
					fbError := fbGripper.fbError;
					ePortalState := E_PortalState_New.eError;		
				END_IF
			END_IF
		END_IF
		
	E_PortalState_New.eSetJob:
		HMI.bAllJobsSend := FALSE;
		IF bReady THEN
			//Weiterer Auftrag in Auftragsreihenfolge
			IF nCntActiveJobs >= 1 AND aJobBuffer[0].eJobType = E_JobType.E_JobType_NewStone THEN 
				aJobBuffer[0].fStartPosX := stActJob.fDestPosX;
				aJobBuffer[0].fStartPosY := stActJob.fDestPosY;
				stActJob := aJobBuffer[0];
				
				eTargetPortalState := E_PortalState_New.eMoveToStone;
				ePortalState := E_PortalState_New.eDebug;
				fSetJobHeight := STONE_POS_FIELD_Z + STONE_HEIGHT;
				
				//ipNcCtrl.M_NewJob(stActJob.fStartPosX, stActJob.fStartPosY, STONE_POS_FIELD_Z + STONE_HEIGHT);
				//ePortalState := E_PortalState_New.eMoveToStone;
			//Weiterer Auftrag in Auftragsreihenfolge
			ELSIF nCntActiveJobs >= 1 AND aJobBuffer[0].eJobType = E_JobType.E_JobType_RemoveStone THEN 
				aJobBuffer[0].fStartPosX := stActJob.fDestPosX;
				aJobBuffer[0].fStartPosY := stActJob.fDestPosY;
				stActJob := aJobBuffer[0];
				
				eTargetPortalState := E_PortalState_New.eMoveToStone;
				ePortalState := E_PortalState_New.eDebug;
				fSetJobHeight := STONE_POS_FIELD_Z; 
				
				//ipNcCtrl.M_NewJob(stActJob.fStartPosX, stActJob.fStartPosY, STONE_POS_FIELD_Z);
				//ePortalState := E_PortalState_New.eMoveToStone;
			END_IF
		ELSE
			nStateJobSelect := M_SetJob_New();
			CASE nStateJobSelect OF
				-1: ePortalState := E_PortalState_New.eEStop;
				0: bReady := FALSE;
				1: bReady := TRUE;
					//Mehr als ein gleichzeitiger Auftrag (NewStone)
					IF nCntActiveJobs >= 1 AND aJobBuffer[0].eJobType = E_JobType.E_JobType_NewStone THEN		
						stActJob := aJobBuffer[0];
						//ipNcCtrl.M_NewJob(stActJob.fStartPosX, stActJob.fStartPosY, fStonePosZFromMag);
						//ePortalState := E_PortalState_New.eMoveToStone;
						fSetJobHeight := fStonePosZFromMag;
						eTargetPortalState := E_PortalState_New.eMoveToStone;
						ePortalState := E_PortalState_New.eDebug;
					//Mehr als ein gleichzeitiger Auftrag (RemoveStone)
					ELSIF nCntActiveJobs >= 1 AND aJobBuffer[0].eJobType = E_JobType.E_JobType_RemoveStone THEN
						stActJob := aJobBuffer[0];
						//ipNcCtrl.M_NewJob(stActJob.fStartPosX, stActJob.fStartPosY, STONE_POS_FIELD_Z);
						//ePortalState := e_PortalState_New.eMoveToStone;
						fSetJobHeight := STONE_POS_FIELD_Z;
						eTargetPortalState := E_PortalState_New.eMoveToStone;
						ePortalState := E_PortalState_New.eDebug;
					//Normaler MoveStone-Auftrag
					ELSIF nCntActiveJobs <= -1 THEN	
						stActJob := aJobBuffer[0];
						ipNcCtrl.M_NewJob(stActJob.fStartPosX, stActJob.fStartPosY, STONE_POS_FIELD_Z);
						ePortalState := E_PortalState_New.eMoveToStone;
					ELSE
						ipNcCtrl.M_NewJob(HMI.fPortalPosIdleX, HMI.fPortalPosIdleY, HMI.fPortalPosIdleZ);
						ePortalState := E_PortalState_New.eHome; //oder Error???
					END_IF
			END_CASE
		END_IF
			
	E_PortalState_New.eDebug:
		IF NOT ipNcCtrl.P_Busy THEN
			ipNcCtrl.M_NewJob(stActJob.fStartPosX, stActJob.fStartPosY, fSetJobHeight);
			ePortalState := eTargetPortalState;
		END_IF
	
	E_PortalState_New.eMoveToStone:
		IF NOT ipNcCtrl.P_Busy THEN 				//Warten bis Position erreicht
			IF ipNcCtrl.P_Error THEN				//Error
				fbError.M_Set(1, 'Achsenfehler', ePortalState, eID := ipNcCtrl.P_ErrID, eSrc := ipNcCtrl.P_ErrSrc);
				ePortalState := E_PortalState_New.eError;
			ELSE
				eTargetPortalState := E_PortalState_New.eTrspStone;
				ePortalState := E_PortalState_New.eCloseGripper;
			END_IF 
		END_IF
		
	E_PortalState_New.eCloseGripper:
		fbGripper(bEnable := TRUE, bClose := TRUE, bOpen := FALSE);
		IF NOT fbGripper.bBusy AND fbGripper.bGripperClosed THEN
			IF NOT fbGripper.fbError.bError THEN
				fbGripper(bClose := FALSE);
				IF fbGripper.bStoneInGripper THEN //Stein von Teilesensor erkannt
					IF stActJob.eJobType = E_JobType_NewStone THEN //Stein aus Magazin entnommen
						IF NOT bStampReset THEN
							aMagCounter[nSelectedMag] := aMagCounter[nSelectedMag] - 1;
						ELSE
							bStampReset := FALSE;
						END_IF
						ipNcCtrl.M_NewJob(stActJob.fDestPosX, stActJob.fDestPosY, STONE_POS_FIELD_Z); 
					ELSIF stActJob.eJobType = E_JobType.E_JobType_RemoveStone AND nCntActiveJobs > 1 AND aJobBuffer[1].fStartPosX <> 0 AND aJobBuffer[1].fStartPosY <> 0 THEN
						stActJob.fDestPosX := aJobBuffer[1].fStartPosX;
						stActJob.fDestPosY := aJobBuffer[1].fStartPosY;
						ipNcCtrl.M_NewJob(stActJob.fDestPosX, stActJob.fDestPosY, STONE_POS_FIELD_Z + STONE_HEIGHT);
					ELSIF (stActJob.eJobType = E_JobType.E_JobType_RemoveStone AND nCntActiveJobs = 1) OR (stActJob.eJobType = E_JobType.E_JobType_RemoveStone AND aJobBuffer[1].fStartPosX <> 0 AND aJobBuffer[1].fStartPosY <> 0) THEN
						stActJob.fDestPosX := STACK_POS_X;
						stActJob.fDestPosY := aMagYPositions[nSelectedMag];
						ipNcCtrl.M_NewJob(stActJob.fDestPosX, stActJob.fDestPosY, STACK_POS_Z_BASE_REMOVE + (nPosInMag-1)*STONE_HEIGHT);
					ELSIF stActJob.eJobType =  E_JobType.E_JobType_MoveStone THEN
						ipNcCtrl.M_NewJob(stActJob.fDestPosX, stActJob.fDestPosY, STONE_POS_FIELD_Z); 
					END_IF
					ePortalState := eTargetPortalState;					
				ELSE
					fbError.M_Set(1804, 'Keinen Stein gegriffen!', ePortalState, eID := E_ErrorIDs.eNoStoneInGripper, eSrc := E_ErrorSrcs.eGripper);
					fbGripper(bOpen := TRUE);
					IF aJobBuffer[0].nJobID = 0 THEN
						ePortalState := E_PortalState_New.eIdle;
					ELSE
						bReady := FALSE;
						ePortalState := E_PortalState_New.eSetJob;
					END_IF
				END_IF
			ELSE
				fbError := fbGripper.fbError;
				ePortalState := E_PortalState_New.eError;
			END_IF
		END_IF
	
	E_PortalState_New.eTrspStone:
		IF NOT ipNcCtrl.P_Busy THEN
			IF ipNcCtrl.P_Error THEN
				fbError.M_Set(1, 'Achsenfehler', ePortalState, eID := ipNcCtrl.P_ErrID, eSrc := ipNcCtrl.P_ErrSrc);
				ePortalState := E_PortalState_New.eError;
			ELSE
				ePortalState := E_PortalState_New.eOpenGripper;
			END_IF 
		END_IF
		
	E_PortalState_New.eError:
		// TODO: Was passiert hier???
	
	E_PortalState_New.eStampTriggered:
		IF NOT ipNcCtrl.P_Busy THEN 
			IF ipNcCtrl.P_Error THEN 	
				fbError.M_Set(1, 'Achsfehler', ePortalState, eID := ipNcCtrl.P_ErrID, eSrc := ipNcCtrl.P_ErrSrc);
				ePortalState := E_PortalState_New.eError;
			ELSE
				fbError.M_Set(1, 'Federung ausgelöst', ePortalState, eID := E_ErrorIDs.eStamp, eSrc := E_ErrorSrcs.ePortal);
				IF aJobBuffer[0].nJobID <> 0 AND aJobBuffer[0].eJobType = E_JobType.E_JobType_RemoveStone THEN
					ePortalState := E_PortalState_New.eSetJob;
				ELSIF aJobBuffer[0].nJobID = 0 THEN
					ePortalState := E_PortalState_New.eIdle;
				ELSIF aJobBuffer[0].nJobID <> 0 AND aJobBuffer[0].eJobType = E_JobType.E_JobType_MoveStone THEN
					ipNcCtrl.M_NewJob(fTargetPosX := aAxis[X].NcToPlc.ActPos, fTargetPosY := aAxis[Y].NcToPlc.ActPos, fTargetPosZ := aAxis[Z].NcToPlc.ActPos+ 10);
					eTargetPortalState := E_PortalState_New.eTrspStone;
				ELSIF aJobBuffer[0].nJobID <> 0 AND aJobBuffer[0].eJobType = E_JobType.E_JobType_NewStone THEN
					ePortalState := E_PortalState_New.eSetJob; //TODO: testen?
				END_IF
			END_IF 
		ELSE
			ipNcCtrl.M_CancleJob();
		END_IF
		
	E_PortalState_New.eHome:
		IF NOT ipNcCtrl.P_Busy THEN
			IF ipNcCtrl.P_Error THEN
				fbError.M_Set(1, 'Achsenfehler', ePortalState, eID := ipNcCtrl.P_ErrID, eSrc := ipNcCtrl.P_ErrSrc);
				ePortalState := E_PortalState_New.eError;
			ELSE
				fbAxesEnable.M_DisableAxes();
				ePortalState := E_PortalState_New.eIdle;
			END_IF 
		END_IF
		
	E_PortalState_New.eManualMode:
		A_CollsionAvoidance();
		fbGripper(bEnable := TRUE, bClose := HMI.bCloseGripper, bOpen := HMI.bOpenGripper);
		IF NOT bManualMode THEN
			fbGripper(bEnable := TRUE, bClose := FALSE, bOpen := FALSE);
			fbAxesEnable.M_EnableAxes();
			ipNcCtrl.P_Enable := TRUE;
			IF fbAxesEnable.bAllAxesReady THEN
				ipNcCtrl.M_NewJob(HMI.fPortalPosIdleX, HMI.fPortalPosIdleY, HMI.fPortalPosIdleZ); //Auftrag an Achsen geben: Grundposition anfahren
				ePortalState := E_PortalState_New.eHome;
			END_IF
		END_IF
		
	E_PortalState_New.eEStop:		
		IF NOT ipNcCtrl.P_Busy THEN
			//ipNcCtrl.M_CancleJob();	//TODO: neu testen
			fbAxesEnable.M_DisableAxes();
		END_IF
		IF bSafetyOK THEN
			IF fbError.bError THEN
				ePortalState := E_PortalState_New.eError;
			ELSE
				bCheck := FALSE;
				bCheckedAllMag := FALSE;
				eCheckMagState := E_CheckMagazines_New.eIdle;
				eSetJobState := E_SetJobState.eIdle;;
				nStonesInMag := MAGAZINE_CAPACITY;
				IF M_IsHomed() THEN
					ePortalState := E_PortalState_New.eIdle;
					nCntActiveJobs := 0;		//TODO: Werte hier notwendig/richtig?
					nCntRemoveStones := 0;
					HMI.bAllJobsSend := FALSE;
				ELSE
					ePortalState := E_PortalState_New.eAfterEStop;
					fbAxesEnable.M_EnableAxes();
				END_IF
			END_IF
		END_IF
		
	E_PortalState_New.eAfterEStop:
		fbGripper();
		IF ipNcCtrl.P_ReadyForJob THEN
			nCntActiveJobs := 0;
			nCntRemoveStones := 0;
			eSetJobState := E_SetJobState.eIdle;
			HMI.bAllJobsSend := FALSE;
			IF fbGripper.bGripperClosed AND fbGripper.bStoneInGripper THEN
				stActJob.nJobID := 1;
				stActJob.eJobType := E_JobType_RemoveStone;
				stActJob.bBlack := bLastJobBlack;
				ipNcCtrl.M_NewJob(aAxis[0].NcToPlc.ActPos, aAxis[1].NcToPlc.ActPos, GVL_CONST.STONE_POS_FIELD_Z);
				ePortalState := E_PortalState_New.eTrspStone;
	//TODO: auswählen Stein(e) zurücktransportieren??? Bleibt hier sonst stecken
			ELSE
				ipNcCtrl.M_NewJob(HMI.fPortalPosIdleX, HMI.fPortalPosIdleY, HMI.fPortalPosIdleZ); //Auftrag an Achsen geben: Grundposition anfahren
				ePortalState := E_PortalState_New.eHome;
			END_IF
		END_IF
END_CASE

ACTION A_ClearJobBuffer:
MEMSET(ADR(aJobBuffer), 0, SIZEOF(aJobBuffer));
MEMSET(ADR(stActJob), 0, SIZEOF(stActJob));
nJobCount := 0;
END_ACTION

ACTION A_CollsionAvoidance:
IF aAxis[X].NcToPlc.SetPos < 0 AND aAxis[Z].NcToPlc.SetPos < MIN_MOVE_HEIGHT_Z THEN
	fbAxesEnable.fOverride := HMI.fAxesOverrideMan;
	fbAxesEnable.bEnableXY := FALSE;//erst beide disablen
	fbAxesEnable.bEnableZn := FALSE;
	FOR nMag := 0 TO MAGAZINE_NUMBER - 1 DO
		fbAxesEnable.bEnableZn := fbAxesEnable.bEnableZn OR ABS(aAxis[Y].NcToPlc.SetPos - aMagYPositions[nMag]) < 0.5; //muss über einem der Stapel stehen (Y)
	END_FOR
	fbAxesEnable.bEnableZn := fbAxesEnable.bEnableZn AND ABS(aAxis[X].NcToPlc.SetPos - STACK_POS_X) < 0.5; //muss die X-Position der Stapel haben
	fbAxesEnable.bEnableZn := fbAxesEnable.bEnableZn AND aAxis[Z].NcToPlc.SetPos > 2.4; //Z darf nicht den Boden der Magazine berühren
	IF fbAxesEnable.bEnableZn = FALSE THEN
		FOR nMag := 0 TO MAGAZINE_NUMBER - 1 DO
			fbAxesEnable.bEnableZn := fbAxesEnable.bEnableZn OR ABS(aAxis[Y].NcToPlc.SetPos - aMagYScanPositions[nMag]) < 0.5; //muss über einem der Stapel stehen (Y)
		END_FOR
		fbAxesEnable.bEnableZn := fbAxesEnable.bEnableZn AND ABS(aAxis[X].NcToPlc.SetPos - STACK_SCAN_POS_X) < 0.5; //muss die X-Position der Stapel haben
	END_IF
	fbAxesEnable.bEnableZn := fbAxesEnable.bEnableZn AND NOT fbGripper.bPartSensor;
ELSE
	fbAxesEnable.fOverride := HMI.fAxesOverride;
	IF aAxis[Z].NcToPlc.SetPos > STONE_POS_FIELD_Z + STONE_HEIGHT THEN
		fbAxesEnable.bEnableXY := TRUE;
	ELSE
		fbAxesEnable.bEnableXY := FALSE;
	END_IF
	fbAxesEnable.bEnableZn := TRUE;
END_IF
END_ACTION

ACTION A_Cycle:
fbAxesEnable(stX := aAxis[X], stY := aAxis[Y], stZ := aAxis[Z]);
rTrigStamp(CLK := bStampZAxis);
rTrigCheck(CLK := fbGripper.bPartSensor);

bSafetyErrAck := FALSE;
bQuitEStop := FALSE;

(*SAFETY CHECK*)
IF NOT bSafetyOK AND ePortalState <> E_PortalState_New.eEStop THEN
	fbGripper(bEnable := FALSE, bClose := FALSE, bOpen := FALSE); //Stopp Greifer
	IF ipNcCtrl <> 0 THEN
		ipNcCtrl.P_Enable := FALSE; //Stopp Achsen
	END_IF
	bLastJobBlack := stActJob.bBlack;
	ePortalState := E_PortalState_New.eEStop;
END_IF

IF ipNcCtrl <> 0 THEN
	ipNcCtrl.M_AxisRef(rX := aAxis[X], rY := aAxis[Y], rZ := aAxis[Z]);
	ipNcCtrl.P_bInductiveSensor := fbGripper.bPartSensor;
	ipNcCtrl.M_Cyclic();
END_IF

(*CHECK FOR NEW JOB*)
IF stNewJob.nJobID > 0 AND HMI.bSetJob AND stNewJob.nJobID <> stActJob.nJobID THEN
	IF nJobCount < MAX_JOB_COUNT AND 
		(stNewJob.fStartPosX > 0 AND stNewJob.fStartPosY > 0 OR stNewJob.eJobType = E_JobType_NewStone) AND //Start Pos must be on the display (if not newStone)
		(stNewJob.fDestPosX > 0 AND stNewJob.fDestPosY > 0 OR stNewJob.eJobType = E_JobType_RemoveStone) //End Pos must be on the display (if not removeStone)
	THEN
		IF nJobCount > 0 THEN
			FOR i := 0 TO nJobCount - 1 DO
				IF stNewJob.nJobID = aJobBuffer[i].nJobID THEN
					EXIT;
				END_IF
			END_FOR
			IF i = nJobCount THEN
				aJobBuffer[nJobCount] := stNewJob;
				aJobBuffer[nJobCount].fStartPosX := aJobBuffer[nJobCount].fStartPosX + HMI.fScreenPosOffsetX;
				aJobBuffer[nJobCount].fStartPosY := aJobBuffer[nJobCount].fStartPosY + HMI.fScreenPosOffsetY;
				aJobBuffer[nJobCount].fDestPosX := aJobBuffer[nJobCount].fDestPosX + HMI.fScreenPosOffsetX;
				aJobBuffer[nJobCount].fDestPosY := aJobBuffer[nJobCount].fDestPosY + HMI.fScreenPosOffsetY;
				nJobCount := nJobCount + 1;
			END_IF
		ELSIF nJobCount = 0 THEN
			aJobBuffer[nJobCount] := stNewJob;
			aJobBuffer[nJobCount].fStartPosX := aJobBuffer[nJobCount].fStartPosX + HMI.fScreenPosOffsetX;
			aJobBuffer[nJobCount].fStartPosY := aJobBuffer[nJobCount].fStartPosY + HMI.fScreenPosOffsetY;
			aJobBuffer[nJobCount].fDestPosX := aJobBuffer[nJobCount].fDestPosX + HMI.fScreenPosOffsetX;
			aJobBuffer[nJobCount].fDestPosY := aJobBuffer[nJobCount].fDestPosY + HMI.fScreenPosOffsetY;
			nJobCount := nJobCount + 1;
		END_IF
		HMI.bSetJob := FALSE;
	ELSE
		;//MELDUNG: Kein Platz mehr im Job Buffer
	END_IF
END_IF

fbRTrigSafety(CLK := bSafetyOK);
IF fbRTrigSafety.Q THEN
	FOR i := 0 TO MAGAZINE_NUMBER - 1 DO
		aMagSkipCheck[i] := FALSE;
	END_FOR
	A_ClearJobBuffer();
	IF ipNcCtrl <> 0 THEN
		ipNcCtrl.P_Enable := TRUE;
	END_IF
	bQuit := TRUE;
END_IF

IF ipNcCtrl.P_Error AND ipNcCtrl.P_ErrID = E_ErrorIDs.eNotAllowedDriveDown THEN
	ePortalState := E_PortalState_New.eError;
END_IF

(*RESET/ERROR ACK*)
IF bQuit THEN
	bQuit := FALSE;
	fbAxesEnable.bReset := TRUE;
	bValidateStonePos := FALSE;
	IF fbError.bError THEN
		A_ClearJobBuffer();
		FOR i := 0 TO MAGAZINE_NUMBER - 1 DO
			aMagSkipCheck[i] := FALSE;
		END_FOR
		IF ePortalState = E_PortalState_New.eError THEN
			ePortalState := E_PortalState_New.eAfterEStop;
			fbAxesEnable.M_EnableAxes();
		END_IF
	END_IF
	fbError.M_Reset();
	fbGripper.fbError.M_Reset();
	
	bSafetyErrAck := TRUE;
	bQuitEStop := TRUE;
	
	FOR i := X TO Z DO
		aAxis[i].ReadStatus();
		IF aAxis[i].Status.Error THEN
			fbResetAxis(Axis := aAxis[i], Execute := TRUE);
			fbResetAxis(Axis := aAxis[i], Execute := FALSE);
		END_IF
	END_FOR
	
	IF ipNcCtrl <> 0 THEN
		ipNcCtrl.P_Reset := TRUE;
	END_IF
END_IF

(*SET BUSY*)
bBusy := ePortalState <> E_PortalState_New.eIdle 
	 AND ePortalState <> E_PortalState_New.eError
	 AND ePortalState <> E_PortalState_New.eEStop;
	 
IF rTrigStamp.Q THEN
	IF ipNcCtrl <> 0 THEN
		IF ipNcCtrl.P_Busy THEN
			ipNcCtrl.M_CancleJob();
			ipNcCtrl.M_NewJob(HMI.fPortalPosIdleX, HMI.fPortalPosIdleY, HMI.fPortalPosIdleZ); //Auftrag an Achsen geben: Grundposition anfahren
			ePortalState := E_PortalState_New.eStampTriggered;
		ELSE
			ePortalState := E_PortalState_New.eStampTriggered;
		END_IF
	END_IF
END_IF
END_ACTION

ACTION A_DequeueJob:
IF nJobCount > 0 THEN
	IF nJobCount > 1 THEN
		FOR k := 0 TO nJobCount - 2 DO
			MEMCPY(ADR(aJobBuffer[k]), ADR(aJobBuffer[k + 1]), SIZEOF(aJobBuffer[k]));
		END_FOR
	END_IF
	MEMSET(ADR(aJobBuffer[nJobCount - 1]), 0, SIZEOF(aJobBuffer[nJobCount - 1]));
	nJobCount := nJobCount - 1;
END_IF
END_ACTION

ACTION A_Init:
(*SET INTERFACE*)
ipNcCtrl := fbNciCtrl;

//Fill Arrays	
aMagCounter[0] := MAGAZINE_CAPACITY;
aMagCounter[1] := MAGAZINE_CAPACITY;
aMagCounter[2] := MAGAZINE_CAPACITY;
aMagCounter[3] := MAGAZINE_CAPACITY;
aMagCounter[4] := MAGAZINE_CAPACITY;
aMagCounter[5] := MAGAZINE_CAPACITY;

aMagYPositions[0] := STACK_1_POS_Y;
aMagYPositions[1] := STACK_2_POS_Y;
aMagYPositions[2] := STACK_3_POS_Y;
aMagYPositions[3] := STACK_4_POS_Y;
aMagYPositions[4] := STACK_5_POS_Y;
aMagYPositions[5] := STACK_6_POS_Y;
    
aMagYScanPositions[0] := STACK_1_SCAN_POS_Y;
aMagYScanPositions[1] := STACK_2_SCAN_POS_Y;
aMagYScanPositions[2] := STACK_3_SCAN_POS_Y;
aMagYScanPositions[3] := STACK_4_SCAN_POS_Y;
aMagYScanPositions[4] := STACK_5_SCAN_POS_Y;
aMagYScanPositions[5] := STACK_6_SCAN_POS_Y;
END_ACTION

METHOD M_CheckStoneInMag_New : INT  //0: working; -2: Error; >0 Anzahl Steine in Magazin; -1: keine Steine in Magazin gefunden
VAR_INPUT
	nMagNumber		: INT;
	nPosNumber		: INT;
	

END_VAR
VAR
END_VAR
//Anzahl an Magazinen stimmt nicht überein
IF MAGAZINE_NUMBER <> 6 THEN
	fbError.M_Set(1,'Anzahl festgelegter Magazine falsch!', eCheckMagState, eID := E_ErrorIDs.eInvalidData, eSrc := E_ErrorSrcs.ePlc);
	M_CheckStoneInMag_New := -2;
	RETURN;
END_IF

//Übergebene Steinposition in Magazin ungültig
IF nPosNumber < 1 OR nPosNumber > MAGAZINE_CAPACITY THEN
	fbError.M_Set(1,'Übergebene Steinposition ungültig!', eCheckMagState, eID := E_ErrorIDs.eInvalidData, eSrc := E_ErrorSrcs.ePlc);
	M_CheckStoneInMag_New := -2;
	RETURN;
END_IF

//Übergebene Magazinnummer ungültig
IF nMagNumber <  0 OR nMagNumber >= MAGAZINE_NUMBER THEN
	fbError.M_Set(1,'Übergebene Magazin-Nummer ungültig!', eCheckMagState, eID := E_ErrorIDs.eInvalidData, eSrc := E_ErrorSrcs.ePlc);
	M_CheckStoneInMag_New := -2;
	RETURN;
END_IF

//Gefordertes Magazin muss nicht überprüft werden
IF aMagSkipCheck[nMagNumber] THEN
	IF aMagCounter[nMagNumber] = 0 THEN
		M_CheckStoneInMag_New := -3;
	ELSE
		M_CheckStoneInMag_New := aMagCounter[nMagNumber];
	END_IF
	RETURN;
END_IF

//Steinanzahl im Magazin zu hoch 
IF 
	fbGripper.bPartSensor 
	AND aAxis[Z].NcToPlc.SetPos > STONE_HEIGHT * (MAGAZINE_CAPACITY - 1) + STACK_SCAN_POS_Z_BASE + STONE_HEIGHT*0.8
	AND aAxis[Z].NcToPlc.SetVelo < 0 //abwärtsbewegung
THEN
	fbError.M_Set(1,'Zu viele Steine in Magazin!', ePortalState, eID := E_ErrorIDs.eInvalidData, eSrc := E_ErrorSrcs.ePortal);
	ipNcCtrl.M_CancleJob();
	M_CheckStoneInMag_New := -2;
END_IF


//Suche nach Anzahl Steine im Magazin
CASE eCheckMagState OF 
	E_CheckMagazines_New.eIdle:
		nStonesInMagazin := 4;
		eCheckMagState := E_CheckMagazines_New.eStartNewNCI;
	
	E_CheckMagazines_New.eStartNewNCI:
		ipNcCtrl.M_NewJob(STACK_SCAN_POS_X, aMagYScanPositions[nMagNumber], STACK_POS_Z_BASE + ((nStonesInMagazin-1) * STONE_HEIGHT ));	
		eCheckMagState := E_CheckMagazines_New.eDebug;
		
	E_CheckMagazines_New.eDebug: 
		IF ipNcCtrl.P_Busy THEN
			eCheckMagState := E_CheckMagazines_New.eWaitForPortal;
		END_IF
		
	E_CheckMagazines_New.eWaitForPortal:
		IF rTrigCheck.Q THEN						//Stein gefunden
			aMagCounter[nMagNumber] := nStonesInMagazin;
			M_CheckStoneInMag_New := nStonesInMagazin;
		ELSIF NOT ipNcCtrl.P_Busy AND NOT fbGripper.bPartSensor THEN					
			IF nStonesInMagazin > 1 THEN					//an aktueller Position kein Stein gefunden
				nStonesInMagazin := nStonesInMagazin -1;
				eCheckMagState:= E_CheckMagazines_New.eStartNewNCI;
			ELSE											//gar kein Stein im Magazin gefunden
				aMagCounter[nMagNumber] := 0;
				M_CheckStoneInMag_New := -1;
			END_IF
		END_IF
END_CASE

IF M_CheckStoneInMag_New <> 0 THEN
	aMagSkipCheck[nMagNumber] := TRUE;
	eCheckMagState := E_CheckMagazines_New.eIdle;
END_IF
END_METHOD

METHOD M_IsHomed : BOOL
VAR_INPUT
END_VAR
M_IsHomed := ABS(aAxis[X].NcToPlc.SetPos - HMI.fPortalPosIdleX) < 2
		AND ABS(aAxis[Y].NcToPlc.SetPos - HMI.fPortalPosIdleY) < 2
		AND ABS(aAxis[Z].NcToPlc.SetPos - HMI.fPortalPosIdleZ) < 2;
END_METHOD

METHOD M_SelEmptyPos_New : BOOL
VAR_INPUT
END_VAR
VAR
	bFirstJobBlack : BOOL;
END_VAR
IF aJobBuffer[0].nJobID <> 0 AND aJobBuffer[0].bBlack THEN		//First Job Black or white
	bFirstJobBlack := TRUE;
ELSIF 
	aJobBuffer[0].nJobID <> 0 AND NOT aJobBuffer[0].bBlack THEN
	bFirstJobBlack := FALSE;
END_IF

FOR i := 0 TO (MIN(4,nJobCount) - 1) BY 1 DO		//Suche Anzahl an zum 1. Job gleichfarbigen Job bis max. 4 Jobs
	IF aJobBuffer[i].nJobID <> 0 AND aJobBuffer[i].bBlack = bFirstJobBlack AND aJobBuffer[i].eJobType = E_JobType.E_JobType_RemoveStone THEN
		nCntActiveJobs := nCntActiveJobs + 1;
	ELSE
		EXIT;
	END_IF
END_FOR

WHILE(nCntActiveJobs > 0) DO
	FOR i := SEL(bFirstJobBlack, MAGAZINE_NUMBER/2, 0) TO SEL (bFirstJobBlack, MAGAZINE_NUMBER-1, MAGAZINE_NUMBER/2-1) BY 1 DO //SEL: Entscheide ob schwarze oder weiße Magazine
		IF MAGAZINE_CAPACITY - aMagCounter[i] >= nCntActiveJobs THEN	//genügend freie Plätze in Magazin vorhanden?
			nSelectedMag := i;
			nPosInMag := aMagCounter[i] + 1;	//abzulegende unterste Steinposition (1 ganz unten, 4 ganz oben)
			fStonePosZFromMag := STACK_POS_Z_BASE + STONE_HEIGHT * (nPosInMag - 1);
			nCntRemoveStones := nCntActiveJobs;
			M_SelEmptyPos_New := TRUE;
			EXIT;
		END_IF
	END_FOR
	
	IF M_SelEmptyPos_New THEN
		EXIT;
	END_IF
	IF NOT M_SelEmptyPos_New AND nCntActiveJobs >= 1 THEN
		i := SEL(bFirstJobBlack, MAGAZINE_NUMBER/2, 0);
		nCntActiveJobs := nCntActiveJobs - 1;
	ELSIF NOT M_SelEmptyPos_New AND nCntActiveJobs = 0 THEN
		M_SelEmptyPos_New := FALSE;
		EXIT;
	END_IF
END_WHILE
END_METHOD

METHOD M_SelNewStone_New : BOOL
VAR_INPUT
END_VAR
VAR
	i		: INT;
	j 		: INT;
	bFirstJobBlack	: BOOL;
END_VAR
IF aJobBuffer[0].nJobID <> 0 AND aJobBuffer[0].bBlack THEN		//First Job Black or white
	bFirstJobBlack := TRUE;
ELSIF 
	aJobBuffer[0].nJobID <> 0 AND NOT aJobBuffer[0].bBlack THEN
	bFirstJobBlack := FALSE;
END_IF

FOR i := 0 TO (MIN(4,nJobCount) - 1) BY 1 DO		//Suche Anzahl an zum 1. Job gleichfarbigen Job bis max. 4 Jobs
	IF aJobBuffer[i].nJobID <> 0 AND aJobBuffer[i].bBlack = bFirstJobBlack AND aJobBuffer[i].eJobType = E_JobType.E_JobType_NewStone THEN
		nCntActiveJobs := nCntActiveJobs + 1;
	ELSE
		EXIT;
	END_IF
END_FOR

WHILE(nCntActiveJobs > 0) DO
	FOR i := SEL(bFirstJobBlack, MAGAZINE_NUMBER/2, 0) TO SEL (bFirstJobBlack, MAGAZINE_NUMBER-1, MAGAZINE_NUMBER/2-1) BY 1 DO //SEL: Entscheide ob schwarze oder weiße Magazine
		IF aMagCounter[i] >= nCntActiveJobs THEN	//genügend Steine in einem Magazin vorhanden
			nSelectedMag := i;
			nPosInMag := aMagCounter[i] - nCntActiveJobs + 1;	//zu greifenden Stein (1 ganz unten, 4 ganz oben)
			aJobBuffer[0].fStartPosX := STACK_POS_X;
			aJobBuffer[0].fStartPosY := aMagYPositions[nSelectedMag];
			fStonePosZFromMag := STACK_POS_Z_BASE + STONE_HEIGHT * (nPosInMag - 1);
			M_SelNewStone_New := TRUE;
			EXIT;
		END_IF
	END_FOR
	IF M_SelNewStone_New THEN
		EXIT;
	END_IF
	IF NOT M_SelNewStone_New AND nCntActiveJobs >= 1 THEN
		i := SEL(bFirstJobBlack, MAGAZINE_NUMBER/2, 0);
		nCntActiveJobs := nCntActiveJobs - 1;
	ELSIF NOT M_SelNewStone_New AND nCntActiveJobs = 0 THEN
		//Gar keine Steine gefunden --> TODO: Was jetzt machen???
		M_SelNewStone_New := FALSE;
		EXIT;
	END_IF
END_WHILE
END_METHOD

METHOD M_SetJob_New : INT
VAR_INPUT
END_VAR
VAR
	bTest	: BOOL;
END_VAR
CASE eSetJobState OF 	//TODO: wenn erste mal Fehler bei M_Sel, dann alle aMagSkipCHeck zurücksetzen und neu suchen
	E_SetJobState.eIdle: 
		IF nJobCount > 0 AND aJobBuffer[0].eJobType = E_JobType_MoveStone AND aJobBuffer[0].nJobID <> 0 THEN
			nCntActiveJobs := -1;
			M_SetJob_New := 1;
		ELSIF nJobCount > 0 AND aJobBuffer[0].eJobType = E_JobType_NewStone AND aJobBuffer[0].nJobID <> 0 THEN
			eSetJobState := E_SetJobState.eSelNewStone;
			nCntActiveJobs := 0;
		ELSIF nJobCount > 0 AND aJobBuffer[0].eJobType = E_JobType.E_JobType_RemoveStone AND aJobBuffer[0].nJobID <> 0 THEN
			//IF NOT bCheckedAllMag THEN
			//	FOR i := 0 TO MAGAZINE_NUMBER -1 BY 1 DO
			//		aMagSkipCheck[i] := FALSE;
			//	END_FOR
			//	eSetJobState := E_SetJobState.eCheckAllMagazines;
			//ELSE
			//	eSetJobState := E_SetJobState.eSelRemoveStone;
			//END_IF
			eSetJobState := E_SetJobState.eSelRemoveStone;
			
			nCntActiveJobs := 0;
		ELSIF aJobBuffer[0].nJobID = 0 THEN
			fbError.M_Set(1,'In M_SetJob Auftrag erwartet, aber nicht gefunden!', ePortalState, eID := E_ErrorIDs.eNoJobsFound, eSrc := E_ErrorSrcs.ePortal);
			M_SetJob_New := -1;
		END_IF
		
		nValidationValue := 0;
		nNumChecked := 0;
		
	E_SetJobState.eSelNewStone:
		IF M_SelNewStone_New() THEN
			eSetJobState := E_SetJobState.eValidateNewStone;
		ELSE
			IF bCheckedAllMag THEN
				M_SetJob_New := -1;																	
				fbError.M_Set(1,'Neuer Stein aufnehmen: Keine Steine im Steinlager gefunden!', ePortalState, eID := E_ErrorIDs.eNoStonesFound, eSrc := E_ErrorSrcs.ePortal);
				eSetJobState := E_SetJobState.eIdle;
			ELSE
				FOR i := 0 TO MAGAZINE_NUMBER -1 BY 1 DO
					aMagSkipCheck[i] := FALSE;
				END_FOR
				eSetJobState := E_SetJobState.eCheckAllMagazines;
			END_IF
		END_IF
		
	E_SetJobState.eValidateNewStone:
		nValidationValue := M_CheckStoneInMag_New(nMagNumber := nSelectedMag, nPosNumber := nPosInMag);
		IF nValidationValue = -2 THEN																	//direkter Fehler
			eSetJobState := E_SetJobState.eIdle;
			M_SetJob_New := -1;
		ELSIF nValidationValue > 0 AND nValidationValue-nCntActiveJobs+1 = nPosInMag THEN				//Gefundenes Magazin korrekt
			eSetJobState := E_SetJobState.eIdle;
			M_SetJob_New := 1;
		ELSIF nValidationValue = -1 OR (nValidationValue > 0 AND nValidationValue <> nPosInMag) OR nValidationValue = -3 THEN 
			//TODO TESTEN: ?? kein Stein in Magazin gefunden oder Anzahl stimmen nicht überein??
			//--> Problem Endlos-Schleife?
			IF bCheckedAllMag THEN 
				M_SetJob_New := -1;
				fbError.M_Set(1,'Beim Aufbauen kein Stein in Magazin gefunden!', ePortalState, eID := E_ErrorIDs.eNoStonesFound, eSrc := E_ErrorSrcs.ePortal);
				eSetJobState := E_SetJobState.eIdle;
			ELSE
				FOR i := 0 TO MAGAZINE_NUMBER -1 BY 1 DO
					aMagSkipCheck[i] := FALSE;
				END_FOR
				eSetJobState := E_SetJobState.eCheckAllMagazines;
			END_IF
		END_IF
		
		IF nValidationValue <> 0 AND eSetJobState <> E_SetJobState.eCheckAllMagazines THEN
			eSetJobState := E_SetJobState.eIdle;
		END_IF
		
	E_SetJobState.eSelRemoveStone:
		IF M_SelEmptyPos_New() THEN
			eSetJobState := E_SetJobState.eValidateRemoveStone;
		ELSE
			IF bCheckedAllMag THEN 
				M_SetJob_New := -1;
				fbError.M_Set(1,'Beim Abräumen keine freien Steinlager gefunden!', ePortalState, eID := E_ErrorIDs.eClearFieldNoCapacityFound, eSrc := E_ErrorSrcs.ePortal);
				eSetJobState := E_SetJobState.eIdle;
			ELSE
				FOR i := 0 TO MAGAZINE_NUMBER -1 BY 1 DO
					aMagSkipCheck[i] := FALSE;
				END_FOR
				eSetJobState := E_SetJobState.eCheckAllMagazines;
			END_IF
		END_IF
		
	E_SetJobState.eValidateRemoveStone:
		nValidationValue := M_CheckStoneInMag_New(nMagNumber := nSelectedMag, nPosNumber := nPosInMag);
		IF nValidationValue = -2 THEN	
			M_SetJob_New := -1;
		ELSIF nValidationValue > 0 AND nValidationValue + 1 = nPosInMag THEN	//Gefundenes Magazin korrekt mit bis zu drei Steinen Platz
			M_SetJob_New := 1;
		ELSIF nValidationValue = -3 AND nValidationValue + 4 = nPosInMag THEN	//Überprüfung geskippt,  mit 4 Steinen Platz
			M_SetJob_New := 1;
		ELSIF nValidationValue = -1 THEN										//Gefundenes Magazin korrekt mit 4 Steinen Platz
			nPosInMag := 1;
			fStonePosZFromMag := STACK_POS_Z_BASE;
			M_SetJob_New := 1;
		ELSIF nValidationValue = 0 THEN
			bTest := TRUE;
		ELSE //TESTEN: Anzahl stimmen nicht überein--> TODO: jetzt M_SelNewStone_New() neu durchlaufen lassen, nMag[] ist schon in Methode auf 0 gesetzt
			IF bCheckedAllMag THEN
				M_SetJob_New := -1;
				fbError.M_Set(1,'Beim Abräumen keine freien Steinlager gefunden!', ePortalState, eID := E_ErrorIDs.eClearFieldNoCapacityFound, eSrc := E_ErrorSrcs.ePortal);
				eSetJobState := E_SetJobState.eIdle;
			ELSE
				eSetJobState := E_SetJobState.eSelRemoveStone;
			END_IF
		END_IF
		
		IF nValidationValue <> 0 AND eSetJobState <> E_SetJobState.eSelRemoveStone THEN
			eSetJobState := E_SetJobState.eIdle;
		END_IF
		
	E_SetJobState.eCheckAllMagazines:
		IF aMagSkipCheck[nNumChecked] THEN
			nNumChecked := nNumChecked + 1;
		ELSE
			nValidationValue := M_CheckStoneInMag_New(nMagNumber := nNumChecked, nPosNumber := 1);
		END_IF
		IF nValidationValue >= 1 OR nValidationValue = -1 OR nValidationValue = -3 THEN
			IF nNumChecked = MAGAZINE_NUMBER-1 THEN
				bCheckedAllMag := TRUE;
				nNumChecked := 0;
				IF nJobCount > 0 AND aJobBuffer[0].eJobType = E_JobType.E_JobType_RemoveStone AND aJobBuffer[0].nJobID <> 0 THEN
					eSetJobState := E_SetJobState.eSelRemoveStone;
				ELSIF nJobCount > 0 AND aJobBuffer[0].eJobType = E_JobType_NewStone AND aJobBuffer[0].nJobID <> 0 THEN
					eSetJobState := E_SetJobState.eSelNewStone;
				END_IF
			ELSE
				nValidationValue := 0;
				nNumChecked := nNumChecked + 1;
			END_IF
		END_IF
	
	E_SetJobState.eAxesNotReady:
		IF fbAxesEnable.bAllAxesReady THEN
			eSetJobState := E_SetJobState.eIdle;
		END_IF
END_CASE

IF NOT fbAxesEnable.bAllAxesReady THEN
	eSetJobState := E_SetJobState.eAxesNotReady;
END_IF
END_METHOD

END_FUNCTION_BLOCK

// ---- POUs/Aktorik/FB_Gripper.TcPOU
FUNCTION_BLOCK FB_Gripper
VAR_INPUT
	bEnable:					BOOL;
	bClose:						BOOL;
	bOpen:						BOOL;
END_VAR                     	
VAR_OUTPUT                  	
	fbError:					FB_Error;	
	bStoneInGripper:			BOOL;
	bPartSensor			AT %I*:	BOOL;
	bBusy:						BOOL;	
END_VAR                     	
VAR CONSTANT                	
	GRIPPER_MOVE_TIME:			TIME := T#120MS;
	GRIPPER_TIMEOUT:			TIME := T#300MS;
END_VAR
VAR
	eState:						E_GripperState;
	bGripperOpen:				BOOL; //kein Sensor
	bGripperClosed:				BOOL; //kein Sensor
	bGripperFullClosed	AT %I*:	BOOL;	
	bOpenGripper		AT %Q*:	BOOL;	
	bCloseGripper		AT %Q*:	BOOL;
	fbTimer:					TON := (PT := GRIPPER_TIMEOUT);
	
(* ******** SIMULATION ************* *)	
	fbTimerSimu:				TON := (PT := GRIPPER_MOVE_TIME);
END_VAR

CASE eState OF
(* ******** INITIALISIERUNG ************* *)	
	E_GripperState_INIT:
		IF bGripperClosed THEN
			eState := E_GripperState_CLOSED;
		ELSIF bGripperOpen THEN
			eState := E_GripperState_OPENED;
		ELSE
			eState := E_GripperState_UNDEFINED;
		END_IF
		
(* ******** GREIFER ÖFFNET ************* *)		
	E_GripperState_OPENING:
		IF NOT bEnable THEN
			bOpenGripper := FALSE;
			eState := E_GripperState_UNDEFINED;
		ELSIF NOT bClose AND bOpen THEN
			IF bGripperOpen THEN
				bOpenGripper := FALSE;
				eState := E_GripperState_OPENED;
				fbError.M_Reset();
			END_IF
		ELSIF NOT bClose AND NOT bOpen OR bClose AND bOpen THEN
			bOpenGripper := FALSE;
			eState := E_GripperState_UNDEFINED;
		ELSIF bClose AND NOT bOpen THEN
			bOpenGripper := FALSE;
			bCloseGripper := TRUE;
			eState := E_GripperState_CLOSING;
		END_IF
		
(* ******** GREIFER OFFEN ************* *)	
	E_GripperState_OPENED:
		IF bClose AND NOT bOpen THEN
			bCloseGripper := TRUE;
			eState := E_GripperState_CLOSING;
		END_IF
		
(* ******** GREIFER SCHLIEßT ************* *)	
	E_GripperState_CLOSING:
		IF NOT bEnable THEN
			bCloseGripper := FALSE;
			eState := E_GripperState_UNDEFINED;
		ELSIF bClose AND NOT bOpen THEN
			IF bGripperClosed THEN
				eState := E_GripperState_CLOSED;
				fbError.M_Reset();
			END_IF
		ELSIF NOT bClose AND NOT bOpen OR bClose AND bOpen THEN
			bCloseGripper := FALSE;
			eState := E_GripperState_UNDEFINED;
		ELSIF NOT bClose AND bOpen THEN
			bCloseGripper := FALSE;
			bOpenGripper := TRUE;
			eState := E_GripperState_OPENING;
		END_IF
		
(* ******** GREIFER GESCHLOSSEN ************* *)	
	E_GripperState_CLOSED:
		IF bOpen AND NOT bClose THEN
			bCloseGripper := FALSE;
			bOpenGripper := TRUE;
			eState := E_GripperState_OPENING;
		END_IF
		
(* ******** GREIFER POSITION UNDEFINIERT ************* *)	
	E_GripperState_UNDEFINED: //Position zwischen den Endlagen
		IF bClose AND NOT bOpen AND NOT bGripperClosed THEN
			bCloseGripper := TRUE;
			eState := E_GripperState_CLOSING;
		END_IF
		IF bOpen AND NOT bClose AND NOT bGripperOpen THEN
			bOpenGripper := TRUE;
			eState := E_GripperState_OPENING;
		END_IF

END_CASE

bBusy := eState = E_GripperState_CLOSING OR eState = E_GripperState_OPENING;

(* ******** TIMEOUT CHECK ************* *)	
fbTimer(IN := eState = E_GripperState_OPENING
			OR eState = E_GripperState_CLOSING);
IF fbTimer.Q THEN
	IF eState = E_GripperState_OPENING THEN
		fbError.M_Set(1817, 'Greifer erreicht Endposition beim Oeffnen nicht!', eState, eID := E_ErrorIDs.eTimeout, eSrc := E_ErrorSrcs.eGripper);
	ELSIF eState = E_GripperState_CLOSING THEN
		fbError.M_Set(1817, 'Greifer erreicht Endposition beim Schliessen nicht!', eState, eID := E_ErrorIDs.eTimeout, eSrc := E_ErrorSrcs.eGripper);
	END_IF
END_IF

(* ******** OUTPUT CHECK ************* *)
IF bGripperClosed AND bGripperOpen
	OR bOpenGripper AND bCloseGripper THEN
	fbError.M_Set(1798, 'Ungültige IO Daten', eState, eID := E_ErrorIDs.eInvalidData, eSrc := E_ErrorSrcs.eGripper);
END_IF

(* ******** SIMULATION ************* *)	
fbTimerSimu(IN := eState = E_GripperState_OPENING OR eState = E_GripperState_CLOSING);
IF bGripperFullClosed THEN
	bStoneInGripper := FALSE;
	bGripperClosed := TRUE;
ELSIF fbTimerSimu.Q THEN
	IF eState = E_GripperState_OPENING THEN
		bGripperClosed := FALSE;
		bStoneInGripper := FALSE;
		bGripperOpen := TRUE;
	END_IF
	IF eState = E_GripperState_CLOSING THEN
		bStoneInGripper := TRUE;
		bGripperOpen := FALSE;
		bGripperClosed := TRUE;
	END_IF
ELSE
	IF eState <> E_GripperState_CLOSED THEN
		bGripperClosed := FALSE;
		bStoneInGripper := FALSE;
	END_IF
	IF eState <> E_GripperState_OPENED THEN
		bGripperOpen := FALSE;
	END_IF
END_IF

END_FUNCTION_BLOCK

// ---- POUs/Aktorik/FB_AxesEnable.TcPOU
FUNCTION_BLOCK FB_AxesEnable
VAR_INPUT
	bEnableAxes: 		BOOL := TRUE;
	bEnableXY:			BOOL;
	bEnableZp:			BOOL;
	bEnableZn:			BOOL;
	bReset:				BOOL;
	fOverride:			LREAL := 10;
END_VAR             	
VAR_OUTPUT          	
	bAllAxesReady:		BOOL := FALSE;
	fbError:			FB_Error;
END_VAR             	
VAR_IN_OUT          	
	stX:				AXIS_REF;
	stY:				AXIS_REF;
	stZ:				AXIS_REF;
END_VAR
VAR	
//Freigaben
	fbPowerX:			MC_Power;
	fbPowerY:			MC_Power;
	fbPowerZ:			MC_Power;
END_VAR


IF NOT (__ISVALIDREF(stX) AND __ISVALIDREF(stY) AND __ISVALIDREF(stZ)) THEN
	fbError.M_Set(1798, 'Üngültige Referenz der Achsen', 0, eID := E_ErrorIDs.eInvalidReference, eSrc := E_ErrorSrcs.ePlc);
	RETURN;
END_IF

IF bReset THEN
	fbError.M_Reset();
	bReset := FALSE;
END_IF

stX.ReadStatus();
stY.ReadStatus();
stZ.ReadStatus();

fbPowerX(
	Enable:=bEnableAxes AND bEnableXY, 
	Enable_Positive:=bEnableAxes AND bEnableXY, 
	Enable_Negative:=bEnableAxes AND bEnableXY, 
	Override:=fOverride, 
	BufferMode:= , 
	Axis:=stX, 
	Status=> , 
	Busy=> , 
	Active=> , 
	Error=> , 
	ErrorID=> );
	
fbPowerY(
	Enable:=bEnableAxes AND bEnableXY, 
	Enable_Positive:=bEnableAxes AND bEnableXY, 
	Enable_Negative:=bEnableAxes AND bEnableXY, 
	Override:=fOverride, 
	BufferMode:= , 
	Axis:=stY, 
	Status=> , 
	Busy=> , 
	Active=> , 
	Error=> , 
	ErrorID=> );	
	
fbPowerZ(
	Enable:=bEnableAxes, 
	Enable_Positive:=bEnableAxes AND bEnableZp, 
	Enable_Negative:=bEnableAxes AND bEnableZn, 
	Override:=fOverride, 
	BufferMode:= , 
	Axis:=stZ, 
	Status=> , 
	Busy=> , 
	Active=> , 
	Error=> , 
	ErrorID=> );		
	
bAllAxesReady := stX.Status.Operational AND stY.Status.Operational AND stZ.Status.Operational;
IF fbPowerX.Error THEN
	fbError.M_Set(fbPowerX.ErrorID, 'Achse X Error', 0, eID := E_ErrorIDs.eAxisRelease, eSrc := E_ErrorSrcs.eAxisX);
ELSIF fbPowerY.Error THEN
	fbError.M_Set(fbPowerY.ErrorID, 'Achse Y Error', 0, eID := E_ErrorIDs.eAxisRelease, eSrc := E_ErrorSrcs.eAxisY);
ELSIF fbPowerZ.Error THEN
	fbError.M_Set(fbPowerZ.ErrorID, 'Achse Z Error', 0, eID := E_ErrorIDs.eAxisRelease, eSrc := E_ErrorSrcs.eAxisZ);
END_IF

METHOD M_DisableAxes
VAR_INPUT
END_VAR
bEnableAxes:= FALSE;
bEnableXY:= FALSE;
bEnableZp:= FALSE; 
bEnableZn:= FALSE;
END_METHOD

METHOD M_EnableAxes
VAR_INPUT
END_VAR
bEnableAxes:= TRUE;
bEnableXY:= TRUE;
bEnableZp:= TRUE; 
bEnableZn:= TRUE;
END_METHOD

END_FUNCTION_BLOCK

// ---- POUs/Aktorik/FB_NciCtrl.TcPOU
FUNCTION_BLOCK FB_NciCtrl IMPLEMENTS I_NC_Ctrl
VAR CONSTANT
	stEmptyCommand:		ST_PositionCmd := (nNo:=0, fPosX:=0, fPosY:=0, fPosZ:=0, fVelo:=0, bExact := FALSE);
END_VAR
VAR
	VELO:				LREAL := 2000;
	DEBUG_RATIO:		LREAL := 0.3;
	bEnable:			BOOL;
	bReset:				BOOL;
	bBusy:				BOOL;
	fbError:			FB_Error;
	eState:				E_NCI_STATE;
	
	rAxisX:				REFERENCE TO AXIS_REF;
	rAxisY:				REFERENCE TO AXIS_REF;
	rAxisZ:				REFERENCE TO AXIS_REF;
	
	fTargetX:			LREAL;
	fTargetY:			LREAL;
	fTargetZ:			LREAL;
	
	fNextTargetX:		LREAL;
	fNextTargetY:		LREAL;
	fNextTargetZ:		LREAL;
	
//NCI	
	stItpToPlc AT %I*:	NcToPlc_NciChannel_Ref;
	stPlcToItp AT %Q*:	PLCTONC_NCICHANNEL_REF;
	
	nFilledRows: 		INT	:= 0;
	nCounter: 			INT	:= 0;
	
	nCommands:			UINT;
	aPositionCmds: 		ARRAY[0..3] OF ST_PositionCmd;	
	
	fbBuildGroup:		CfgBuildExt3DGroup;
	fbClearGroup:		CfgReconfigGroup;
	
	fbFeedTablePrep:	FB_NciFeedTablePreparation;	(* fb that is good for the preparation of the table - inserts elements to table *)
	fbFeedTable: 		FB_NciFeedTable;	(* is responsible that the prepared table is transfered to nc-kernel *)
	
	fbNciEStop:			ItpEStopEx;
	fbNciReset:			ItpResetEx2;
	bEStop:				BOOL;
	
	stNciFeedTable:		ST_NciFeedGroupTable;	(* table that holds the entries *)
	
	stGeoStart: 		ST_NciGeoStart;		(* structure for starting pos - required if first entry is a circle *)
	stGeoLine: 			ST_NciGeoLine;		(* structure for straight line segment *)
	stVertexSmoothing: 	ST_NciVertexSmoothing;	(* structure to enable blending of serveral geo entries *)
	stEndOfTables: 		ST_NciEndOfTables;	(* structure to indicate end of tables *)	
END_VAR
VAR
	bInductiveSensor: BOOL;
	nCntForAxesReady: UINT := 0;
END_VAR

CASE eState OF
	E_NCI_State_INIT:
		IF __ISVALIDREF(rAxisX) AND __ISVALIDREF(rAxisY) AND __ISVALIDREF(rAxisZ) THEN		
			eState := E_NCI_State_IDLE;
			nCntForAxesReady := 0;
		END_IF
		
	E_NCI_State_IDLE:
		M_AxesReady();
		IF fTargetX <> fNextTargetX OR fTargetY <> fNextTargetY OR fTargetZ <> fNextTargetZ THEN
			IF M_AxesReady() (*AND nCntForAxesReady < 5*) THEN
				IF bInductiveSensor 
					AND fNextTargetZ < rAxisZ.NcToPlc.ActPos 
					AND fNextTargetX - 3 > rAxisX.NcToPlc.ActPos AND fNextTargetX + 3 < rAxisX.NcToPlc.ActPos
					AND fNextTargetY - 3 > rAxisY.NcToPlc.ActPos AND fNextTargetY + 3 < rAxisX.NcToPlc.ActPos
				THEN
					fbError.M_Set(1, 'Neuer NCI-Auftrag: tiefer fahren nicht erlaubt', eState, E_ErrorIDs.eNotAllowedDriveDown, E_ErrorSrcs.eAxisCtrlNci);
					eState	:= E_NCI_State_ERROR;
				ELSE
					fTargetX := fNextTargetX;
					fTargetY := fNextTargetY;
					fTargetZ := fNextTargetZ;
					eState := E_NCI_State_BUILD_GROUP;
					bReset := FALSE;
					bBusy := TRUE;
					nCntForAxesReady := 0;
				END_IF
			(*ELSIF NOT M_AxesReady() AND nCntForAxesReady < 5 THEN
				nCntForAxesReady := nCntForAxesReady + 1;*)
			ELSE
				fbError.M_Set(1, 'Achsen nicht betriebsbereit', eState, E_ErrorIDs.eAxesNotReady, E_ErrorSrcs.eAxisCtrlNci);
			END_IF
		END_IF
		
	E_NCI_State_BUILD_GROUP://Interpolationsgruppe bauen 		
		fbBuildGroup(
			bExecute:=TRUE, 
			nGroupId:=ItpGetGroupId(sNciToPlc:=stItpToPlc) , 
			nXAxisId:=rAxisX.NcToPlc.AxisId, 
			nYAxisId:=rAxisY.NcToPlc.AxisId, 
			nZAxisId:=rAxisZ.NcToPlc.AxisId, 
			nQ1AxisId:= 0, 
			nQ2AxisId:= 0, 
			nQ3AxisId:= 0, 
			nQ4AxisId:= 0, 
			nQ5AxisId:= 0);
			
		IF NOT fbBuildGroup.bBusy THEN
			IF NOT fbBuildGroup.bErr THEN
				ItpSetOverridePercent(HMI.fAxesOverride, stPlcToItp);
				A_PrepareTable();
				eState	:= E_NCI_State_FEED_TABLE;
			ELSE
				fbError.M_Set(fbBuildGroup.nErrId, 'Fehler beim Bauen der Gruppe!', eState, eID := E_ErrorIDs.eBuildGroup, eSrc := E_ErrorSrcs.eAxisCtrlNci);
				eState	:= E_NCI_State_ERROR;
			END_IF
			fbBuildGroup(bExecute:=FALSE); 
		END_IF
		
	E_NCI_State_FEED_TABLE: //Tabelle füllen
		fbFeedTable(
			bExecute:=TRUE,
			bReset:=FALSE,
			bLogFeederEntries:=FALSE,
			stFeedGroupTable:=stNciFeedTable,
			stNciToPlc:=stItpToPlc);
		IF fbFeedTable.bFeedingDone THEN //Alle Befehle sind in Tabelle gespeichert
			eState	:= E_NCI_State_RUN;
		ELSIF fbFeedTable.bError THEN
			fbError.M_Set(fbFeedTable.nErrorId, 'Fehler beim Tabelle füllen', eState, eID := E_ErrorIDs.eFillTable, eSrc := E_ErrorSrcs.eAxisCtrlNci);
			eState := E_NCI_State_CLEAR_GROUP;
		END_IF
		
	E_NCI_State_RUN:
		IF NOT bEnable THEN
			eState := E_NCI_State_ABORT;
		ELSE
			fbFeedTable(stFeedGroupTable:=stNciFeedTable, stNciToPlc:=stItpToPlc);
			IF fbFeedTable.bChannelDone THEN //Bewegung abgeschlossen
				fbFeedTable(bExecute:=FALSE, bReset:=FALSE, stFeedGroupTable:=stNciFeedTable, stNciToPlc:=stItpToPlc);
				eState := E_NCI_State_CLEAR_GROUP;
			ELSIF fbFeedTable.bError THEN
				fbError.M_Set(fbFeedTable.nErrorId, 'Fehler beim Fahren des Kommandos', eState, eID := E_ErrorIDs.eAbsMove, eSrc := E_ErrorSrcs.eAxisCtrlNci);
				eState := E_NCI_State_CLEAR_GROUP;
			END_IF
		END_IF

	E_NCI_State_ABORT:
		fbFeedTable(bExecute := FALSE, stFeedGroupTable:=stNciFeedTable, stNciToPlc:=stItpToPlc);
		fbNciEStop(sNciToPlc := stItpToPlc);
		IF NOT fbNciEStop.bBusy THEN
			IF NOT fbNciEStop.bErr THEN
				fbFeedTablePrep(bResetTable:=TRUE, stFeedGroupTable:=stNciFeedTable);
				fbFeedTablePrep(bResetTable:=FALSE, stFeedGroupTable:=stNciFeedTable);
			ELSE
				fbError.M_Set(fbNciEStop.nErrId, 'Fehler beim EStop!', eState, eID := E_ErrorIDs.eStopAxis, eSrc := E_ErrorSrcs.eAxisCtrlNci);
			END_IF
			bEStop := TRUE;
			eState := E_NCI_State_CLEAR_GROUP;
			fbNciEStop(sNciToPlc := stItpToPlc, bExecute := FALSE);
		END_IF
	
	E_NCI_State_CLEAR_GROUP:
		fbClearGroup(bExecute := TRUE, nGroupId := stItpToPlc.GrpId);
		IF NOT fbClearGroup.bBusy THEN
			fbClearGroup(bExecute := FALSE, nGroupId := stItpToPlc.GrpId);
			IF NOT fbError.bError THEN
				IF NOT fbClearGroup.bErr THEN
					IF bEStop THEN
						bEStop := FALSE;
						eState := E_NCI_State_ESTOP;
					ELSE			
						eState := E_NCI_State_IDLE;
					END_IF
				ELSE
					fbError.M_Set(fbClearGroup.nErrId, 'Fehler beim Auflösen der Gruppe!', eState, eID := E_ErrorIDs.eClearGroup, eSrc := E_ErrorSrcs.eAxisCtrlNci);
					eState := E_NCI_State_ERROR;
				END_IF
			ELSE
				eState := E_NCI_State_ERROR;
			END_IF
		END_IF
	
	E_NCI_State_ESTOP:
		IF bReset THEN
			fbFeedTable(bExecute := TRUE, bReset := TRUE, stFeedGroupTable := stNciFeedTable, stNciToPlc := stItpToPlc);
			IF NOT fbFeedTable.bResetBusy THEN
				IF NOT fbFeedTable.bError THEN
					fbFeedTable(bExecute := FALSE, bReset := FALSE, stFeedGroupTable := stNciFeedTable, stNciToPlc := stItpToPlc);
					bReset := FALSE;
					nCntForAxesReady := 0;
					eState := E_NCI_State_IDLE;
				ELSE
					fbError.M_Set(fbFeedTable.nErrorId, 'Fehler beim Tabellen-Reset!', eState, eID := E_ErrorIDs.eReset, eSrc := E_ErrorSrcs.eAxisCtrlNci);
					eState := E_NCI_State_ERROR;
				END_IF
			END_IF
		END_IF
	
	E_NCI_State_ERROR:
		IF bReset THEN
			fbFeedTable(bExecute := TRUE, bReset := TRUE, stFeedGroupTable := stNciFeedTable, stNciToPlc := stItpToPlc);
			IF NOT fbFeedTable.bResetBusy THEN
				IF NOT fbFeedTable.bError THEN
					fbFeedTable(bExecute := FALSE, bReset := FALSE, stFeedGroupTable := stNciFeedTable, stNciToPlc := stItpToPlc);
					bReset := FALSE;
					nCntForAxesReady := 0;
					eState := E_NCI_State_IDLE;
					fbError.M_Reset();
				END_IF
			END_IF
		END_IF
END_CASE

ACTION A_PrepareTable:
(* clear all old entries & reset to default data *)
fbFeedTablePrep(
	bResetAll:=TRUE,
	stFeedGroupTable:=stNciFeedTable );

(* fill up table with start position *)
stGeoStart.fPosX	:= rAxisX.NcToPlc.SetPos;
stGeoStart.fPosY	:= rAxisY.NcToPlc.SetPos;
stGeoStart.fPosZ	:= rAxisZ.NcToPlc.SetPos;
fbFeedTablePrep(
	nEntryType:= E_NciEntryTypeGeoStart,
	pEntry:= ADR(stGeoStart) ,
	bResetAll:=FALSE,
	bResetTable:= FALSE,
	stFeedGroupTable:= stNciFeedTable,
	nFilledRows=>nFilledRows);
IF fbFeedTablePrep.bError THEN
	IF fbFeedTablePrep.nErrorId = ErrNciFeedTableFull THEN
		fbError.M_Set(fbFeedTablePrep.nErrorId, 'Tabelle voll!', eState, eID := E_ErrorIDs.eFillTable, eSrc := E_ErrorSrcs.eAxisCtrlNci);
		eState := E_NCI_State_ERROR;
	ELSE
		fbError.M_Set(fbFeedTablePrep.nErrorId, 'Fehler beim Tabelle speisen!', eState, eID := E_ErrorIDs.eFillTable, eSrc := E_ErrorSrcs.eAxisCtrlNci);
		eState := E_NCI_State_ERROR;
	END_IF
	RETURN;
END_IF


(* enable vertex smoothing *)
stVertexSmoothing.fRadius	:= 50.0; 	(* max. blending radius *)
stVertexSmoothing.nDisplayIndex	:= 0;
stVertexSmoothing.nType	:= 2; (* type: parabola *)
stVertexSmoothing.nSubtype	:= 3; (* adapative tolerance radius *)
fbFeedTablePrep(
	nEntryType:= E_NciEntryTypeVertexSmoothing,
	pEntry:= ADR(stVertexSmoothing) ,
	bResetTable:= FALSE,
	stFeedGroupTable:= stNciFeedTable,
	nFilledRows=>nFilledRows);
IF fbFeedTablePrep.bError THEN
	IF fbFeedTablePrep.nErrorId = ErrNciFeedTableFull THEN
		fbError.M_Set(fbFeedTablePrep.nErrorId, 'Tabelle voll!', eState, eID := E_ErrorIDs.eFillTable, eSrc := E_ErrorSrcs.eAxisCtrlNci);
		eState := E_NCI_State_ERROR;
	ELSE
		fbError.M_Set(fbFeedTablePrep.nErrorId, 'Fehler beim Tabelle speisen!', eState, eID := E_ErrorIDs.eFillTable, eSrc := E_ErrorSrcs.eAxisCtrlNci);
		eState := E_NCI_State_ERROR;
	END_IF
	RETURN;
END_IF

A_SetPosCommands();

(* add positions of the array to the feeder table *)
FOR nCounter := 0 TO TO_INT(nCommands) - 1 DO
	stGeoLine.nDisplayIndex	:= aPositionCmds[nCounter].nNo;
	stGeoLine.fEndPosX		:= aPositionCmds[nCounter].fPosX;
	stGeoLine.fEndPosY		:= aPositionCmds[nCounter].fPosY;
	stGeoLine.fEndPosZ		:= aPositionCmds[nCounter].fPosZ;
	stGeoLine.fVelo			:= aPositionCmds[nCounter].fVelo; (*mm per sec*)
	stGeoLine.bAccurateStop := aPositionCmds[nCounter].bExact; 
	fbFeedTablePrep(
		nEntryType:= E_NciEntryTypeGeoLine,
		pEntry:= ADR(stGeoLine),
		bResetTable:= FALSE,
		stFeedGroupTable:= stNciFeedTable,
		nFilledRows=>nFilledRows);
	IF fbFeedTablePrep.bError THEN
		IF fbFeedTablePrep.nErrorId = ErrNciFeedTableFull THEN
			fbError.M_Set(fbFeedTablePrep.nErrorId, 'Tabelle voll!', eState, eID := E_ErrorIDs.eFillTable, eSrc := E_ErrorSrcs.eAxisCtrlNci);
			eState := E_NCI_State_ERROR;
		ELSE
			fbError.M_Set(fbFeedTablePrep.nErrorId, 'Fehler beim Tabelle speisen!', eState, eID := E_ErrorIDs.eFillTable, eSrc := E_ErrorSrcs.eAxisCtrlNci);
			eState := E_NCI_State_ERROR;
		END_IF
		RETURN;
	END_IF
END_FOR

(* add end of tables flag *)
fbFeedTablePrep(
	nEntryType:= E_NciEntryTypeEndOfTables,
	pEntry:= ADR(stEndOfTables) ,
	bResetTable:= FALSE,
	stFeedGroupTable:= stNciFeedTable,
	nFilledRows=>nFilledRows);
IF fbFeedTablePrep.bError THEN
	IF fbFeedTablePrep.nErrorId = ErrNciFeedTableFull THEN
		fbError.M_Set(fbFeedTablePrep.nErrorId, 'Tabelle voll!', eState, eID := E_ErrorIDs.eFillTable, eSrc := E_ErrorSrcs.eAxisCtrlNci);
		eState := E_NCI_State_ERROR;
	ELSE
		fbError.M_Set(fbFeedTablePrep.nErrorId, 'Fehler beim Tabelle speisen!', eState, eID := E_ErrorIDs.eFillTable, eSrc := E_ErrorSrcs.eAxisCtrlNci);
		eState := E_NCI_State_ERROR;
	END_IF
	RETURN;
END_IF
END_ACTION

ACTION A_SetPosCommands:
FOR nCounter := 0 TO 3 DO
	aPositionCmds[nCounter] := stEmptyCommand;
END_FOR
nCommands := 0;

IF rAxisZ.NcToPlc.SetPos < MIN_MOVE_HEIGHT_Z AND (ABS(fTargetX - rAxisX.NcToPlc.SetPos) > 2 OR ABS(fTargetY - rAxisY.NcToPlc.SetPos) > 2) THEN
	aPositionCmds[nCommands].nNo   := 10*(nCommands + 1);
	aPositionCmds[nCommands].fPosX := rAxisX.NcToPlc.SetPos;
	aPositionCmds[nCommands].fPosY := rAxisY.NcToPlc.SetPos;
	aPositionCmds[nCommands].fPosZ := MIN_MOVE_HEIGHT_Z; //erst vertikal Gefahrenbereich verlassen, dann zum Ziel fahren
	aPositionCmds[nCommands].fVelo := VELO;
	aPositionCmds[nCommands].bExact := FALSE;
	nCommands := nCommands + 1;
END_IF
aPositionCmds[nCommands].nNo   := 10*(nCommands + 1);	
aPositionCmds[nCommands].fPosX := fTargetX;
aPositionCmds[nCommands].fPosY := fTargetY;
aPositionCmds[nCommands].fVelo := VELO;
IF fTargetZ < MIN_MOVE_HEIGHT_Z AND (ABS(fTargetX - rAxisX.NcToPlc.SetPos) > 2 OR ABS(fTargetY - rAxisY.NcToPlc.SetPos) > 2) THEN
	aPositionCmds[nCommands].fPosZ := MIN_MOVE_HEIGHT_Z;
ELSE
	aPositionCmds[nCommands].fPosZ := fTargetZ;
	IF fTargetZ < MIN_MOVE_HEIGHT_Z THEN
		aPositionCmds[nCommands].fVelo := VELO * DEBUG_RATIO;
	END_IF
END_IF
aPositionCmds[nCommands].bExact := FALSE;
nCommands := nCommands + 1;

IF aPositionCmds[nCommands - 1].fPosZ <> fTargetZ THEN
	aPositionCmds[nCommands].nNo   := 10*(nCommands + 1);
	aPositionCmds[nCommands].fPosX := fTargetX;
	aPositionCmds[nCommands].fPosY := fTargetY;
	aPositionCmds[nCommands].fPosZ := fTargetZ; 
	aPositionCmds[nCommands].fVelo := VELO * DEBUG_RATIO;
	aPositionCmds[nCommands].bExact := FALSE;
	nCommands := nCommands + 1;
END_IF
END_ACTION

METHOD M_AxesReady : BOOL
VAR_INPUT
END_VAR
IF __ISVALIDREF(rAxisX) AND __ISVALIDREF(rAxisY) AND __ISVALIDREF(rAxisZ) THEN		
	rAxisX.ReadStatus();
	rAxisY.ReadStatus();
	rAxisZ.ReadStatus();
	IF rAxisX.Status.Operational AND rAxisY.Status.Operational AND rAxisZ.Status.Operational THEN
		M_AxesReady := TRUE;
	END_IF
END_IF
END_METHOD

METHOD M_AxisRef
VAR_INPUT
	rX	: REFERENCE TO AXIS_REF;
	rY	: REFERENCE TO AXIS_REF;
	rZ	: REFERENCE TO AXIS_REF;
END_VAR

rAxisX REF= rX;
rAxisY REF= rY;
rAxisZ REF= rZ;
END_METHOD

METHOD M_CancleJob
IF eState = E_NCI_State_RUN THEN
	eState := E_NCI_State_ABORT;
	bReset := TRUE;
END_IF
END_METHOD

METHOD M_Cyclic
THIS^();

bBusy := eState <> E_NCI_State_IDLE
	 AND eState <> E_NCI_State_ERROR
	 AND eState <> E_NCI_State_ESTOP;
	
IF bReset THEN
	fTargetX := 0;
	fTargetY := 0;
	fTargetZ := 0;
	
	fNextTargetX := 0;
	fNextTargetY := 0;
	fNextTargetZ := 0;
END_IF
END_METHOD

METHOD M_NewJob
VAR_INPUT
	fTargetPosX	: LREAL;
	fTargetPosY	: LREAL;
	fTargetPosZ	: LREAL;
END_VAR
VAR
	bTest	: BOOL;
END_VAR
IF(fTargetPosX < 1 AND fTargetPosX > -1) AND (fTargetPosY < 1 AND fTargetPosY > -1) THEN
	bTest := TRUE;
END_IF
fNextTargetX := fTargetPosX;
fNextTargetY := fTargetPosY;
fNextTargetZ := fTargetPosZ;
END_METHOD

PROPERTY P_bInductiveSensor : BOOL
SET
bInductiveSensor := P_bInductiveSensor;
END_SET
END_PROPERTY

PROPERTY P_Busy : BOOL
GET
P_Busy := bBusy;
END_GET
END_PROPERTY

PROPERTY P_Enable : BOOL
SET
bEnable := P_Enable;
END_SET
END_PROPERTY

PROPERTY P_ErrID : E_ErrorIDs
GET
P_ErrID := fbError.eErrorID;
END_GET
END_PROPERTY

PROPERTY P_Error : BOOL
GET
P_Error := fbError.bError;
END_GET
END_PROPERTY

PROPERTY P_ErrSrc : E_ErrorSrcs
GET
P_ErrSrc := fbError.eErrorSrc;
END_GET
END_PROPERTY

{warning 'add property implementation'}
PROPERTY P_ReadyForJob : BOOL
GET
P_ReadyForJob := eState = E_NCI_State_IDLE AND M_AxesReady();
END_GET
END_PROPERTY


PROPERTY P_Reset : BOOL
SET
bReset := P_Reset;
END_SET
END_PROPERTY

END_FUNCTION_BLOCK

// ---- POUs/Safety/FB_SafetyMonitoring.TcPOU
FUNCTION_BLOCK FB_SafetyMonitoring
VAR_INPUT
END_VAR
VAR_OUTPUT
	bQuitDone:				BOOL;
	fbError:				FB_Error;
	
	bLightCurtainOk AT %I*:	BOOL;
	bEStopButtonOk 	AT %I*:	BOOL;
END_VAR
VAR
	fbGroup:				FB_SafeGroup;

	fbMonLightCurtain:		FB_SafeMon;
	fbMonEStop:				FB_SafeMon;
	fbMonSafetyGroup:		FB_SafeMon;
	fbEStop:				FB_SafeEStop;
	
	nDrvInfoData1	AT %I*:	WORD;
	nDrvInfoData2	AT %I*:	WORD;
	nDrvInfoData3	AT %I*:	WORD;
	bCollectEDM		AT %Q*:	BOOL;
END_VAR

fbGroup(bIsReset => bQuitDone);
fbMonLightCurtain();
fbMonEStop();
fbMonSafetyGroup();
fbEStop();
IF fbMonLightCurtain.fbError.bError 
	OR fbMonEStop.fbError.bError
	OR fbMonSafetyGroup.fbError.bError
	OR fbEStop.fbError.bError
	OR fbGroup.fbError.bError
THEN
	fbError.M_Set(1, 'Safety-Fehler', 0, E_ErrorIDs.eUndefinedError, E_ErrorSrcs.eSafety);
END_IF

bCollectEDM := NOT nDrvInfoData1.8
			AND NOT nDrvInfoData2.8
			AND NOT nDrvInfoData3.8;
			
IF NOT bEStopButtonOk THEN
	fbError.M_Set(1, 'Not-Aus betätigt', 0, E_ErrorIDs.eEStopPressed, eSrc := E_ErrorSrcs.eSafety);
ELSIF NOT bLightCurtainOk THEN
	fbError.M_Set(1, 'Lichtgitter ausgelöst', 0, E_ErrorIDs.eLightCurtain, eSrc := E_ErrorSrcs.eSafety);
ELSIF fbError.bError THEN
	fbError.M_Reset();
END_IF

END_FUNCTION_BLOCK

// ---- POUs/Safety/FB_SafeGroup.TcPOU
FUNCTION_BLOCK FB_SafeGroup
VAR_INPUT
END_VAR
VAR_OUTPUT
	bIsReset:		BOOL;
	fbError:		FB_Error;
END_VAR
VAR
	nDiag	AT %I*:	USINT;
	nState	AT %I*:	USINT;
	sMsg:			STRING;
	i:				INT;
END_VAR

bIsReset := nState = 5;
CASE nState OF
	0: //undefined
		IF NOT fbError.bError THEN
			fbError.M_Set(1, 'Undefinierter State!', nState, eID := E_ErrorIDs.eUndefinedState, eSrc := E_ErrorSrcs.eSafetyGroup);
		END_IF
	1: //RUN
		IF fbError.bError THEN
			fbError.M_Reset();
		END_IF
	2:;
	4://Error
		CASE nDiag OF
			0:
				fbError.M_Set(1, 'Ungültiger Wert!', nDiag, eID := E_ErrorIDs.eInvalidData, eSrc := E_ErrorSrcs.eSafetyGroup); //nState sagt Error, nDiag sagt aber kein Error! 
			1:	
				fbError.M_Set(1, 'Safety FB Error!', nDiag, eID := E_ErrorIDs.eSafetyFbError, eSrc := E_ErrorSrcs.eSafetyGroup); 
			2:	
				fbError.M_Set(1, 'Safety Kommunikationsfehler!', nDiag, eID := E_ErrorIDs.eCommError, eSrc := E_ErrorSrcs.eSafetyGroup); 
			3:	
				fbError.M_Set(1, 'Module Fault!', nDiag, eID := E_ErrorIDs.eModuleFault, eSrc := E_ErrorSrcs.eSafetyGroup); 
			4:	
				fbError.M_Set(1, 'Vergleich-Fehler!', nDiag, eID := E_ErrorIDs.eCompareError, eSrc := E_ErrorSrcs.eSafetyGroup); 
			5:	                                              
				fbError.M_Set(1, 'Timeout Com-Fehler!', nDiag, eID := E_ErrorIDs.eTimeout, eSrc := E_ErrorSrcs.eSafetyGroup);
			6:	                                              
				fbError.M_Set(1, 'Restart Fehler!', nDiag, eID := E_ErrorIDs.eReset, eSrc := E_ErrorSrcs.eSafetyGroup); 
			ELSE                                              
				fbError.M_Set(1, 'Ungültiger Wert!', nDiag, eID := E_ErrorIDs.eInvalidData, eSrc := E_ErrorSrcs.eSafetyGroup);
		END_CASE
	5,6,7,16,17:;
	ELSE //undefined
		IF NOT fbError.bError THEN
			fbError.M_Set(1, 'Undefinierter State!', nState, eID := E_ErrorIDs.eUndefinedState, eSrc := E_ErrorSrcs.eSafetyGroup);
		END_IF
END_CASE

END_FUNCTION_BLOCK

// ---- POUs/Safety/FB_SafeMon.TcPOU
FUNCTION_BLOCK FB_SafeMon
VAR_INPUT
END_VAR
VAR_OUTPUT
	bSafeState:		BOOL;
	bIsReset:		BOOL;
	fbError:		FB_Error;
END_VAR
VAR
	{attribute 'displaymode':='binary'}
	nDiag	AT %I*:	UINT;
	nState	AT %I*:	USINT;
	sMsg:			STRING;
	i:				INT;
END_VAR

bSafeState := nState = 3;
bIsReset := nState = 5;
CASE nState OF
	0: //undefined
		IF NOT fbError.bError THEN
			fbError.M_Set(1, 'Undefinierter State!', nState, eID := E_ErrorIDs.eUndefinedState, eSrc := E_ErrorSrcs.eSafetyFb);
		END_IF
	1: //RUN
		IF fbError.bError THEN
			fbError.M_Reset();
		END_IF
	2:;
	3:;
	4://Error
		IF NOT fbError.bError THEN
			IF nDiag.0 THEN
				sMsg := CONCAT(sMsg, 'DiskrepGr1,');
			END_IF
			IF nDiag.1 THEN
				sMsg := CONCAT(sMsg, 'DiskrepGr2,');
			END_IF
			IF nDiag.2 THEN
				sMsg := CONCAT(sMsg, 'DiskrepGr3,');
			END_IF
			IF nDiag.3 THEN
				sMsg := CONCAT(sMsg, 'DiskrepGr4,');
			END_IF
			IF nDiag.4 THEN
				sMsg := CONCAT(sMsg, 'EDM1,');
			END_IF
			IF nDiag.5 THEN
				sMsg := CONCAT(sMsg, 'EDM2,');
			END_IF
			IF nDiag.8 THEN
				sMsg := CONCAT(sMsg, 'DiskrepErrGr1Plus');
			END_IF
			IF nDiag.9 THEN
				sMsg := CONCAT(sMsg, 'DiskrepErrGr2Plus');
			END_IF
			IF nDiag.10 THEN
				sMsg := CONCAT(sMsg, 'DiskrepErrGr3Plus');
			END_IF
			IF nDiag.11 THEN
				sMsg := CONCAT(sMsg, 'DiskrepErrGr4Plus');
			END_IF
			
			fbError.M_Set(1, sMsg, TO_INT(nDiag), eID := E_ErrorIDs.eSafetyFbError, eSrc := E_ErrorSrcs.eSafetyFb);
		END_IF
	5,6,8:;
	ELSE //undefined
		IF NOT fbError.bError THEN
			fbError.M_Set(1, 'Undefinierter State!', nState, eID := E_ErrorIDs.eUndefinedState, eSrc := E_ErrorSrcs.eSafetyFb);
		END_IF
END_CASE

END_FUNCTION_BLOCK

// ---- POUs/Safety/FB_SafeEStop.TcPOU
FUNCTION_BLOCK FB_SafeEStop
VAR_INPUT
END_VAR
VAR_OUTPUT
	bSafeState:		BOOL;
	bIsReset:		BOOL;
	fbError:		FB_Error;
END_VAR
VAR
	{attribute 'displaymode':='binary'}
	nDiag	AT %I*:	UINT;
	nState	AT %I*:	USINT;
	sMsg:			STRING;
	i:				INT;
END_VAR

bSafeState := nState = 3;
bIsReset := nState = 5;
CASE nState OF
	0: //undefined
		IF NOT fbError.bError THEN
			fbError.M_Set(1, 'Undefinierter State!', nState, eID := E_ErrorIDs.eUndefinedState, eSrc := E_ErrorSrcs.eSafetyFb);
		END_IF
	1: //RUN
		IF fbError.bError THEN
			fbError.M_Reset();
		END_IF
	2:;
	3:;
	4://Error
		IF NOT fbError.bError THEN
			IF nDiag.0 THEN
				sMsg := CONCAT(sMsg, 'DiskrepGr1,');
			END_IF
			IF nDiag.1 THEN
				sMsg := CONCAT(sMsg, 'DiskrepGr2,');
			END_IF
			IF nDiag.2 THEN
				sMsg := CONCAT(sMsg, 'DiskrepGrSec,');
			END_IF
			IF nDiag.4 THEN
				sMsg := CONCAT(sMsg, 'EDM1,');
			END_IF
			IF nDiag.5 THEN
				sMsg := CONCAT(sMsg, 'EDM2,');
			END_IF
			IF nDiag.8 THEN
				sMsg := CONCAT(sMsg, 'DiskrepErrGr1Plus');
			END_IF
			IF nDiag.9 THEN
				sMsg := CONCAT(sMsg, 'DiskrepErrGr2Plus');
			END_IF
			IF nDiag.10 THEN
				sMsg := CONCAT(sMsg, 'DiskrepErrSecPlus');
			END_IF
			
			fbError.M_Set(1, sMsg, TO_INT(nDiag), eID := E_ErrorIDs.eSafetyFbError, eSrc := E_ErrorSrcs.eSafetyFb);
		END_IF
	5,6,7,8,9:;
	ELSE //undefined
		IF NOT fbError.bError THEN
			fbError.M_Set(1, 'Undefinierter State!', nState, eID := E_ErrorIDs.eUndefinedState, eSrc := E_ErrorSrcs.eSafetyFb);
		END_IF
END_CASE

END_FUNCTION_BLOCK

// ---- POUs/Zeug/FB_FuseControl.TcPOU
FUNCTION_BLOCK FB_FuseControl
VAR_INPUT
	bResetChannels:	BOOL;
END_VAR
VAR_OUTPUT
	fbError:		FB_Error;
END_VAR
VAR
	fbBlockFuse:	FB_BlockEconomySmart;
	nChannel:		INT;
END_VAR

fbBlockFuse();
FOR nChannel := fbBlockFuse.MIN_CHANNEL TO fbBlockFuse.MAX_CHANNEL DO
	CASE fbBlockFuse.Status[nChannel] OF 
		fbBlockFuse.STATUS_TRIP:
			fbError.M_Set(1, CONCAT('Sicherung hat ausgelöst! Kanal ', TO_STRING(nChannel)), 0, E_ErrorIDs.eFuseTripped, E_ErrorSrcs.eFuse);
			EXIT;
		fbBlockFuse.STATUS_OVERCURRENT:
			fbError.M_Set(1, CONCAT('Sicherung Überstrom! Kanal ', TO_STRING(nChannel)), 0, E_ErrorIDs.eFuseOvercurrent, E_ErrorSrcs.eFuse);
			EXIT;
		fbBlockFuse.STATUS_OFF:
			fbError.M_Set(1, CONCAT('Sicherung ausgeschaltet! Kanal ', TO_STRING(nChannel)), 0, E_ErrorIDs.eFuseOff, E_ErrorSrcs.eFuse);
			EXIT;
		fbBlockFuse.STATUS_ON:
			IF fbError.bError THEN
				fbError.M_Reset();				
			END_IF
		ELSE
			fbError.M_Set(1, CONCAT('Sicherung ausgeschaltet! Kanal ', TO_STRING(nChannel)), 0, E_ErrorIDs.eFuseOff, E_ErrorSrcs.eFuse);
			EXIT;
	END_CASE
END_FOR

IF fbBlockFuse.FuseTripped AND bResetChannels THEN
	fbBlockFuse.reset();
END_IF

END_FUNCTION_BLOCK

// ---- POUs/Zeug/FB_BlockEconomySmart.TcPOU
//Block Economy Smart 
//FB is able to control and read all values from Block Ecomemy Smart Fuse
{attribute 'no_check'}
FUNCTION_BLOCK FB_BlockEconomySmart
VAR CONSTANT 										
	MIN_DATA												:	INT := 0;
	MAX_DATA												:	INT := 90;
//	BASE_CLOCK												:	INT := 120; // MIN: 70 MAX: 200
END_VAR
VAR_OUTPUT CONSTANT
	MIN_CHANNEL												: INT := 1;
	MAX_CHANNEL												: INT := 4;
	STATUS_ON												: BYTE := 0;
	STATUS_OFF												: BYTE := 1;
	STATUS_TRIP												: BYTE := 2;
	STATUS_OVERCURRENT										: BYTE := 3;
END_VAR                         							
VAR_INPUT                       							
	Enable													: BOOL := TRUE; //Enable communication 
	Force													: ARRAY[MIN_CHANNEL..MAX_CHANNEL] OF BOOL; 	// 	simulates channel
	Control													: ARRAY[MIN_CHANNEL..MAX_CHANNEL] OF BOOL; 	// 	Enable/Disable channel 
	SetCtrl													: BOOL := FALSE;		// 	Write channel control to output (Econemy Smart Fuse)
	ResetTrig												: BOOL := FALSE;		// 	Reset tripped fuses/channels
	ReadSetValues											: BOOL := FALSE;		// 	Read trip set value of all cannels 
	ExtProtocolSampleingDivider								: UINT := 0;			//  0 = read only short protocol / >0 = read long protocol every n cycles 					
END_VAR
VAR_OUTPUT
	Voltage													: LREAL;					// [V] actual voltage
	Current													: ARRAY[MIN_CHANNEL..MAX_CHANNEL] OF LREAL;	// [A] actual cannel current[1-8]
	Status													: ARRAY[MIN_CHANNEL..MAX_CHANNEL] OF BYTE;	// Fuse status
	FuseTripped												: BOOL := FALSE;		// min 1 Fuse has tripped
	UpdateCycle												: UINT := 0;			// update Cycle counter
	Busy													: BOOL; 
END_VAR
VAR 
	In												AT%I*	: BOOL;
	Out												AT%Q*	: BOOL;
END_VAR
VAR
//local cache ************************************************************************************
	State													: INT := -1;
	CycleTime												: LREAL; // [ms] Cycle Time of PLC Task
	_BaseClock												: INT := 100; // MIN: 70 MAX: 200
	CurrentCycles											: UDINT;
	CyclePerTick											: UDINT;
	_InternReset											: BOOL;

	BitIdx													: INT;
	SendData												: ARRAY[MIN_DATA..MAX_DATA] OF BOOL;
	Receive													: ARRAY[MIN_DATA..MAX_DATA] OF BOOL;
	
	{attribute 'displaymode':='binary'}
	Temp 													: BYTE;		


				
//trigger *********************************************************************************
	
//timer ***********************************************************************************
	Delay													: TON;
	
//instances ***********************************************************************************             								
	GETCURTASKINDEX											: GETCURTASKINDEX;


//Dummys ****************************************************************************************
	i,j														: INT;
END_VAR

	(* Block Economy Smart communication 					*)
	(********************************************************)

(* Initiat reset of channel ***********************************************)
	IF ResetTrig THEN reset();	END_IF

(* State machine to read and write data ************************************)
	CASE State OF
	-1: // init
		GETCURTASKINDEX();
		CycleTime 											:= TwinCAT_SystemInfoVarList._TaskInfo[GETCURTASKINDEX.index].CycleTime / 10_000;
		IF CycleTime > 0 THEN           						
			CyclePerTick									:= LREAL_TO_UDINT(_BaseClock / CycleTime);	
			CyclePerTick									:= CyclePerTick + (CyclePerTick MOD 2);
			State											:= 0;
		END_IF                          						
																
	0: // idle          
		IF Enable
		THEN    	   
			Busy											:= TRUE; 						
			FOR i := MIN_CHANNEL TO MAX_CHANNEL DO    									
				SendData[i]									:= Control[9-i];
			END_FOR                 						
			SendData[9]										:= SetCtrl;			    	
			SendData[10]									:= extProtocolSampleingDivider <> 0
																AND(	
																(UpdateCycle MOD extProtocolSampleingDivider) = 0
																OR UpdateCycle = 0)
																OR ReadSetValues;
			SendData[11]									:= ReadSetValues;
			BitIdx											:= 0;		
			State											:= SEL(_InternReset, 10, 5); // Reset tripped if flag is true
		ELSE
			Busy											:= FALSE;
			Out												:= FALSE;
			State											:= 0;
			Voltage											:= 0.0;
			MEMSET(ADR(Current),0,SIZEOF(Current));			
			MEMSET(ADR(Status),0,SIZEOF(Status));	        
			FuseTripped										:= FALSE;
			UpdateCycle										:= 0;		
		END_IF
																
	5:	//reset triped          								
		Out													:= TRUE;
		Delay(IN:= NOT Delay.Q, PT := T#600MS);             
															
		IF Delay.Q THEN             						
			_InternReset									:= FALSE;
			Delay(IN := FALSE);                             
			State 											:= 20;
		END_IF                  							
															
	10: // receive	            							
		Out													:= SendData[BitIdx] XOR CurrentCycles <= CyclePerTick / 2;		
															
		IF CurrentCycles >= CyclePerTick					 
		THEN                            	                
			Receive[BitIdx]									:= In;
			CurrentCycles									:= 0;
			BitIdx											:= BitIdx + 1;
			IF BitIdx > 16 AND NOT SendData[10] AND NOT SendData[11]
				OR BitIdx > 89
			THEN
				Out											:= FALSE;
				State										:= 20;
			END_IF                  	
		ELSE	                    	
			CurrentCycles									:= CurrentCycles + 1;
		END_IF
		
	20:	 // interpret
		Delay( IN:= NOT Delay.Q AND NOT IN, PT := TO_TIME(_BaseClock*3));
		IF Delay.Q THEN		// stop Bit		
			Delay(IN := FALSE);
			
